        // Temporary bypass.
        eState := E_IndexState.Complete;


    E_IndexState.WaitingSupportExtended:

        (*
        bSupportExtendRequest := TRUE;

        IF bSupportExtended
            AND bTableReady
            AND bTableLocked
        THEN

            IF bManualMoveActive
                OR bPositionRecoveryActive
            THEN
                eState := E_IndexState.Complete;
            ELSE
                eState := E_IndexState.ProcessPositionReady;
            END_IF

        ELSIF tonStateTimeout.Q THEN

            eFault := E_IndexFault.SupportExtendTimeout;
            eState := E_IndexState.Fault;

        END_IF
        *)

        // Temporary bypass.
        eState := E_IndexState.Complete;


    // =====================================================
    // AUTOMATIC-CYCLE STATES
    // CURRENTLY RETAINED BUT NOT USED BY MANUAL MOVEMENT
    // =====================================================

    E_IndexState.ProcessPositionReady:

        (*
        bSupportExtendRequest := TRUE;
        *)

        IF bReleaseProcessPosition THEN

            bReleaseProcessPosition := FALSE;
            eState := E_IndexState.WaitingOperatorExchange;

        END_IF


    E_IndexState.WaitingOperatorExchange:

        (*
        bSupportExtendRequest := TRUE;
        *)

        IF bOperatorExchangeDone THEN

            bOperatorExchangeDone := FALSE;
            eState := E_IndexState.Complete;

        END_IF


    // =====================================================
    // COMPLETE
    // =====================================================

    E_IndexState.Complete:

        bDonePulse := TRUE;

        bManualMoveActive := FALSE;
        bPositionRecoveryActive := FALSE;
        bWrongPositionSupervisionActive := FALSE;

        eState := E_IndexState.Idle;


    // =====================================================
    // STOPPING
    // =====================================================

    E_IndexState.Stopping:

        // Outputs are already reset at the beginning of this method.
        IF NOT bRotatePortA THEN
            eState := E_IndexState.Idle;
        END_IF


    // =====================================================
    // FAULT
    // =====================================================

    E_IndexState.Fault:

        // No movement outputs are generated while faulted.


END_CASE


// =========================================================
// STATUS MAPPING
// =========================================================

stInternalStatus.eState := eState;
stInternalStatus.eFault := eFault;
stInternalStatus.eCurrentPosition := eCurrentPosition;

stInternalStatus.bReady :=
    eState = E_IndexState.Idle
    OR eState = E_IndexState.ProcessPositionReady;

stInternalStatus.bBusy :=
    // Support states retained for future use.
    (eState = E_IndexState.RetractingSupport)
    OR (eState = E_IndexState.WaitingSupportRetracted)

    OR (eState = E_IndexState.RotatingPortA)
    OR (eState = E_IndexState.WrongPositionRecovery)
    OR (eState = E_IndexState.StoppingPortB)
    OR (eState = E_IndexState.VerifyingPosition)

    // Support states retained for future use.
    OR (eState = E_IndexState.ExtendingSupport)
    OR (eState = E_IndexState.WaitingSupportExtended);

stInternalStatus.bFaulted :=
    eState = E_IndexState.Fault;

stInternalStatus.bDonePulse :=
    bDonePulse;

stInternalStatus.bManualMoveActive :=
    bManualMoveActive;

stInternalStatus.bPositionRecoveryActive :=
    bPositionRecoveryActive;
	
stInternalStatus.bSamePositionDetected :=
    bSamePositionDetected;

stInternalStatus.bWrongPositionTimerActive :=
    bWrongPositionSupervisionActive;

stInternalStatus.bTwoHandRequired :=
    bRequestPending
    OR (
        stInternalStatus.bBusy
        AND NOT bTableLocked
    );

stInternalStatus.bProcessPositionReady :=
    eState = E_IndexState.ProcessPositionReady;

stInternalStatus.bWaitingOperatorExchange :=
    eState = E_IndexState.WaitingOperatorExchange;


// Support feedback remains published for diagnostics, even though it
// is not currently used to permit the movement.
stInternalStatus.bSupportRetracted :=
    bSupportRetracted;

stInternalStatus.bSupportExtended :=
    bSupportExtended;

stInternalStatus.bTableReady :=
    bTableReady;

stInternalStatus.bTableLocked :=
    bTableLocked;
END_METHOD

METHOD PUBLIC GetFault : E_IndexFault
GetFault := eFault;
END_METHOD

METHOD PUBLIC GetState : E_IndexState
GetState := eState;
END_METHOD

METHOD PUBLIC GetStatus : ST_IndexStatus
GetStatus := stInternalStatus;
END_METHOD

METHOD PUBLIC IsDone : BOOL
IsDone := bDonePulse;
END_METHOD

METHOD PUBLIC IsFaulted : BOOL
IsFaulted := eState = E_IndexState.Fault;
END_METHOD

METHOD PUBLIC IsProcessPositionReady : BOOL
IsProcessPositionReady := eState = E_IndexState.ProcessPositionReady;
END_METHOD

METHOD PUBLIC IsReady : BOOL
IsReady := eState = E_IndexState.Idle OR eState = E_IndexState.ProcessPositionReady;
END_METHOD

METHOD PUBLIC ReleaseProcessPosition
IF eState = E_IndexState.ProcessPositionReady THEN bReleaseProcessPosition := TRUE; END_IF
END_METHOD

METHOD PUBLIC RequestManualMove : BOOL
RequestManualMove := FALSE;
IF eState = E_IndexState.Idle AND NOT bRequestPending THEN
    bRequestPending := TRUE;
    bManualMoveActive := TRUE;
    RequestManualMove := TRUE;
END_IF
END_METHOD

METHOD PUBLIC RequestMove : BOOL
RequestMove := FALSE;
IF eState = E_IndexState.Idle AND NOT bRequestPending THEN
    bRequestPending := TRUE;
    bManualMoveActive := FALSE;
    RequestMove := TRUE;
END_IF
END_METHOD

METHOD PUBLIC RequestPositionRecovery : BOOL
RequestPositionRecovery := FALSE;
IF eState = E_IndexState.Idle
   AND NOT bRequestPending
   AND stInternalStatus.eCurrentPosition = E_TablePosition.Unknown
THEN
    bRequestPending := TRUE;
    bManualMoveActive := FALSE;
    bPositionRecoveryActive := TRUE;
    RequestPositionRecovery := TRUE;
END_IF
END_METHOD

METHOD PUBLIC Reset
bRequestPending := FALSE;
bManualMoveActive := FALSE;
bPositionRecoveryActive := FALSE;
bWrongPositionSupervisionActive := FALSE;
bReleaseProcessPosition := FALSE;
bOperatorExchangeDone := FALSE;
eFault := E_IndexFault.None;
eState := E_IndexState.Initialising;
END_METHOD

END_FUNCTION_BLOCK

// ---- POUs/02_Components/Door/FB_MainDoorLock.TcPOU
FUNCTION_BLOCK FB_MainDoorLock
VAR
    eState           : E_MainDoorLockState := E_MainDoorLockState.Disabled;
    eFault           : E_MainDoorLockFault := E_MainDoorLockFault.None;
    stStatusInternal : ST_MainDoorLockStatus;
    tonTransition    : TON;
END_VAR

METHOD PUBLIC Cyclic : BOOL
VAR_INPUT
    bEnableAutomatic       : BOOL;
    bManualEnable          : BOOL;
    bManualLockRequest     : BOOL;
    bManualUnlockRequest   : BOOL;
    bStopRequest           : BOOL;
    bResetRequest          : BOOL;
    bDoorClosed            : BOOL;
    bDoorLocked            : BOOL;
    bIndexBusy             : BOOL;
    bProcessSafePosition   : BOOL;
    tLockTimeout           : TIME;
    tUnlockTimeout         : TIME;
	bDoorUnsafe 		   : BOOL;
END_VAR
VAR_OUTPUT
    bLockOutput            : BOOL;
	
END_VAR
// -----------------------------------------------------------------------------
// Unlock permissive
// -----------------------------------------------------------------------------
stStatusInternal.bUnlockPermissive :=
    NOT bIndexBusy
    AND bProcessSafePosition;


// -----------------------------------------------------------------------------
// This FB only supervises the main door.
//
// The physical locking is performed externally by the pneumatic system and
// TwinSAFE. This FB does not command the door lock.
// -----------------------------------------------------------------------------
bLockOutput := FALSE;


// -----------------------------------------------------------------------------
// Fault reset
// -----------------------------------------------------------------------------
IF bResetRequest THEN

    // The fault cannot be reset while TwinSAFE still reports the door unsafe.
    IF NOT bDoorUnsafe THEN

        eFault := E_MainDoorLockFault.None;

        // Restore the internal state according to the current feedbacks.
        IF bDoorClosed AND bDoorLocked THEN
            eState := E_MainDoorLockState.Locked;
        ELSE
            eState := E_MainDoorLockState.Unlocked;
        END_IF

    END_IF

END_IF


// -----------------------------------------------------------------------------
// Unsafe door condition reported by TwinSAFE
//
// Example:
//     Door not confirmed closed AND lock feedback active.
// -----------------------------------------------------------------------------
IF bDoorUnsafe THEN

    eFault := E_MainDoorLockFault.FeedbackMismatch;
    eState := E_MainDoorLockState.Fault;

END_IF


// -----------------------------------------------------------------------------
// Main door supervision state machine
// -----------------------------------------------------------------------------
CASE eState OF

    // -------------------------------------------------------------------------
    // Disabled
    // -------------------------------------------------------------------------
    E_MainDoorLockState.Disabled:

        IF bEnableAutomatic OR bManualEnable THEN

            IF bDoorClosed
                AND bDoorLocked
                AND NOT bDoorUnsafe
            THEN
                eState := E_MainDoorLockState.Locked;
            ELSE
                eState := E_MainDoorLockState.Unlocked;
            END_IF

        END_IF


    // -------------------------------------------------------------------------
    // Unlocked
    //
    // Wait for the operator to close the door.
    // An open door is not considered a fault in this state.
    // -------------------------------------------------------------------------
    E_MainDoorLockState.Unlocked:

        IF bEnableAutomatic
            OR (bManualEnable AND bManualLockRequest)
        THEN

            IF bDoorClosed AND NOT bDoorUnsafe THEN
                eState := E_MainDoorLockState.Locking;
            END_IF

        END_IF


    // -------------------------------------------------------------------------
    // Locking
    //
    // TwinSAFE and the pneumatic system perform the physical locking.
    // This FB only waits for the safe locked feedback.
    // -------------------------------------------------------------------------
    E_MainDoorLockState.Locking:

        IF bDoorUnsafe THEN

            eFault := E_MainDoorLockFault.FeedbackMismatch;
            eState := E_MainDoorLockState.Fault;

        ELSIF NOT bDoorClosed THEN

            // The door was opened before locking was confirmed.
            // Return to Unlocked without generating a fault.
            eState := E_MainDoorLockState.Unlocked;

        ELSIF bDoorLocked THEN

            eState := E_MainDoorLockState.Locked;

        ELSIF tonTransition.Q THEN

            eFault := E_MainDoorLockFault.LockTimeout;
            eState := E_MainDoorLockState.Fault;

        END_IF


    // -------------------------------------------------------------------------
    // Locked
    // -------------------------------------------------------------------------
    E_MainDoorLockState.Locked:

		// Door feedback inconsistency reported by TwinSAFE.
		IF bDoorUnsafe THEN
	
			eFault := E_MainDoorLockFault.FeedbackMismatch;
			eState := E_MainDoorLockState.Fault;
	
	
		// While automatic locking is required, the door must remain
		// physically closed and locked.
		ELSIF bEnableAutomatic
			AND (
				NOT bDoorClosed
				OR NOT bDoorLocked
			)
		THEN
	
			eFault := E_MainDoorLockFault.FeedbackMismatch;
			eState := E_MainDoorLockState.Fault;
	
	
		// Existing controlled unlock paths remain below.
		ELSIF NOT bEnableAutomatic
			AND bManualEnable
			AND bManualUnlockRequest
			AND stStatusInternal.bUnlockPermissive
		THEN
	
			eState := E_MainDoorLockState.Unlocking;
	
	
		ELSIF NOT bEnableAutomatic
			AND NOT bManualEnable
			AND bStopRequest
			AND stStatusInternal.bUnlockPermissive
		THEN
	
			eState := E_MainDoorLockState.Unlocking;
	
		END_IF


    // -------------------------------------------------------------------------
    // Unlocking
    //
    // The external safety/pneumatic system removes the locking condition.
    // This FB only waits for the lock feedback to disappear.
    // -------------------------------------------------------------------------
    E_MainDoorLockState.Unlocking:

        IF bDoorUnsafe THEN

            eFault := E_MainDoorLockFault.FeedbackMismatch;
            eState := E_MainDoorLockState.Fault;

        ELSIF NOT bDoorLocked THEN

            eState := E_MainDoorLockState.Unlocked;

        ELSIF tonTransition.Q THEN

            eFault := E_MainDoorLockFault.UnlockTimeout;
            eState := E_MainDoorLockState.Fault;

        END_IF


    // -------------------------------------------------------------------------
    // Fault
    // -------------------------------------------------------------------------
    E_MainDoorLockState.Fault:

        // No physical output is controlled by this FB.
        //
        // Recovery requires:
        //   - bDoorUnsafe = FALSE
        //   - bResetRequest = TRUE


    // -------------------------------------------------------------------------
    // Invalid internal state
    // -------------------------------------------------------------------------
    ELSE

        eFault := E_MainDoorLockFault.FeedbackMismatch;
        eState := E_MainDoorLockState.Fault;

END_CASE


// -----------------------------------------------------------------------------
// Transition timer
//
// TwinCAT SEL:
//   G = FALSE -> first value
//   G = TRUE  -> second value
//
// Locking:
//   eState = Locking -> TRUE -> tLockTimeout
//
// Unlocking:
//   eState = Locking -> FALSE -> tUnlockTimeout
// -----------------------------------------------------------------------------
tonTransition(
    IN :=
        (eState = E_MainDoorLockState.Locking)
        OR (eState = E_MainDoorLockState.Unlocking),

    PT := SEL(
        eState = E_MainDoorLockState.Locking,
        tUnlockTimeout,
        tLockTimeout
    )
);

// -----------------------------------------------------------------------------
// Status mapping
// -----------------------------------------------------------------------------
stStatusInternal.eState := eState;
stStatusInternal.eFault := eFault;

stStatusInternal.bDoorClosed := bDoorClosed;
stStatusInternal.bDoorLocked := bDoorLocked;
stStatusInternal.bDoorUnsafe := bDoorUnsafe;


// This indicates that the machine expects the door to be locked.
// It does not command the physical locking mechanism.
stStatusInternal.bLockRequest :=
    bEnableAutomatic
    OR (bManualEnable AND bManualLockRequest);


// Retained only for interface compatibility.
// This FB no longer controls a physical output.
stStatusInternal.bLockOutput := FALSE;


// Door ready for automatic operation
stStatusInternal.bReadyForAutomatic :=
    bEnableAutomatic
    AND bDoorClosed
    AND bDoorLocked
    AND NOT bDoorUnsafe
    AND (eState = E_MainDoorLockState.Locked);


stStatusInternal.bFaulted :=
    eState = E_MainDoorLockState.Fault;


// -----------------------------------------------------------------------------
// Diagnostic message
// -----------------------------------------------------------------------------
IF bDoorUnsafe THEN

    stStatusInternal.sMessage :=
        'Unsafe main door feedback';

ELSE

    CASE eState OF

        E_MainDoorLockState.Disabled:
            stStatusInternal.sMessage :=
                'Main door supervision disabled';

        E_MainDoorLockState.Unlocked:
            stStatusInternal.sMessage :=
                'Waiting for main door to close';

        E_MainDoorLockState.Locking:
            stStatusInternal.sMessage :=
                'Waiting for main door lock feedback';

        E_MainDoorLockState.Locked:
            stStatusInternal.sMessage :=
                'Main door closed and locked';

        E_MainDoorLockState.Unlocking:
            stStatusInternal.sMessage :=
                'Waiting for main door to unlock';

        E_MainDoorLockState.Fault:
            stStatusInternal.sMessage :=
                'Main door supervision fault';

        ELSE
            stStatusInternal.sMessage :=
                'Invalid main door state';

    END_CASE

END_IF


// -----------------------------------------------------------------------------
// Method result
// -----------------------------------------------------------------------------
Cyclic := NOT stStatusInternal.bFaulted;
END_METHOD

METHOD PUBLIC GetStatus : ST_MainDoorLockStatus
GetStatus := stStatusInternal;
END_METHOD

METHOD PUBLIC Initialise
eFault := E_MainDoorLockFault.None;
IF stStatusInternal.bDoorLocked THEN eState := E_MainDoorLockState.Locked; ELSE eState := E_MainDoorLockState.Unlocked; END_IF
tonTransition(IN := FALSE);
END_METHOD

METHOD PUBLIC IsFaulted : BOOL
IsFaulted := stStatusInternal.bFaulted;
END_METHOD

METHOD PUBLIC IsReadyForAutomatic : BOOL
IsReadyForAutomatic := stStatusInternal.bReadyForAutomatic;
END_METHOD

END_FUNCTION_BLOCK

// ---- POUs/02_Components/Index/FB_NestTableManager.TcPOU
FUNCTION_BLOCK FB_NestTableManager
VAR
    aNestInternal           : ARRAY[1..4] OF ST_Nest;
    aNestStatisticsInternal : ARRAY[1..4] OF ST_NestStatistics;
    aPositionToNest         : ARRAY[1..4] OF UINT := [1,2,3,4];
    bInitialised            : BOOL;
    i                       : INT;
    uiNest                  : UINT;
    uiMethodNestId          : UINT;
END_VAR

METHOD PUBLIC ClearOperatorNest
VAR_INPUT ePosition : E_TablePosition; END_VAR
uiMethodNestId := GetNestIdAtPosition(ePosition); IF uiMethodNestId >= 1 AND uiMethodNestId <= 4 THEN aNestInternal[uiMethodNestId].bProcessRequired := FALSE; aNestInternal[uiMethodNestId].bProcessComplete := FALSE; aNestInternal[uiMethodNestId].eDisposition := E_PartDisposition.None; aNestInternal[uiMethodNestId].bDispositionSent := FALSE; aNestInternal[uiMethodNestId].bOperatorExchangeComplete := FALSE; aNestInternal[uiMethodNestId].stPatchDispenseResult.bValid := FALSE; aNestInternal[uiMethodNestId].stHeatStakeResult.bValid := FALSE; aNestInternal[uiMethodNestId].stVisionResult.bValid := FALSE; aNestInternal[uiMethodNestId].stResult.bValid := FALSE; aNestInternal[uiMethodNestId].bStatisticsCounted := FALSE; END_IF
END_METHOD

METHOD PUBLIC Cyclic
VAR_INPUT
    bIndexStable : BOOL;
    eIndexPosition : E_TablePosition;
    eOperatorPosition : E_TablePosition;
    bPartPresent : BOOL;
    aNestEnabled : ARRAY[1..4] OF BOOL;
END_VAR
IF NOT bInitialised THEN
    FOR i := 1 TO 4 DO
        aNestInternal[i].nId := INT_TO_UINT(i);
        aNestStatisticsInternal[i].uiNestId := INT_TO_UINT(i);
    END_FOR
    bInitialised := TRUE;
END_IF
FOR i := 1 TO 4 DO aNestInternal[i].bEnabled := aNestEnabled[i]; END_FOR
IF bIndexStable AND (eIndexPosition <> E_TablePosition.Unknown) THEN
    CASE eIndexPosition OF
        E_TablePosition.Position1:
            aPositionToNest[1] := 1;
            aPositionToNest[2] := 4;
            aPositionToNest[3] := 3;
            aPositionToNest[4] := 2;
        E_TablePosition.Position2:
            aPositionToNest[1] := 2;
            aPositionToNest[2] := 1;
            aPositionToNest[3] := 4;
            aPositionToNest[4] := 3;
        E_TablePosition.Position3:
            aPositionToNest[1] := 3;
            aPositionToNest[2] := 2;
            aPositionToNest[3] := 1;
            aPositionToNest[4] := 4;
        E_TablePosition.Position4:
            aPositionToNest[1] := 4;
            aPositionToNest[2] := 3;
            aPositionToNest[3] := 2;
            aPositionToNest[4] := 1;
    END_CASE
    FOR i := 1 TO 4 DO
        aNestInternal[aPositionToNest[i]].ePosition := UINT_TO_E_TablePosition(INT_TO_UINT(i));
        aNestInternal[i].bPartLoadedPulse := FALSE;
        aNestInternal[i].bPartRemovedPulse := FALSE;
    END_FOR
    uiNest := aPositionToNest[TO_UINT(eOperatorPosition)];
    aNestInternal[uiNest].bPartLoadedPulse := bPartPresent AND NOT aNestInternal[uiNest].bPreviousPartPresent;
    aNestInternal[uiNest].bPartRemovedPulse := NOT bPartPresent AND aNestInternal[uiNest].bPreviousPartPresent;
    aNestInternal[uiNest].bPreviousPartPresent := bPartPresent;
    aNestInternal[uiNest].bPartPresent := bPartPresent;
END_IF
END_METHOD

METHOD PUBLIC GetAllNests : ARRAY[1..4] OF ST_Nest
GetAllNests := aNestInternal;
END_METHOD

METHOD PUBLIC GetAllNestStatistics : ARRAY[1..4] OF ST_NestStatistics
GetAllNestStatistics := aNestStatisticsInternal;
END_METHOD

METHOD PUBLIC GetNestAtPosition : ST_Nest
VAR_INPUT ePosition : E_TablePosition; END_VAR
uiMethodNestId := GetNestIdAtPosition(ePosition); IF uiMethodNestId >= 1 AND uiMethodNestId <= 4 THEN GetNestAtPosition := aNestInternal[uiMethodNestId]; END_IF
END_METHOD

METHOD PUBLIC GetNestIdAtPosition : UINT
VAR_INPUT ePosition : E_TablePosition; END_VAR
IF ePosition >= E_TablePosition.Position1 AND ePosition <= E_TablePosition.Position4 THEN GetNestIdAtPosition := aPositionToNest[TO_UINT(ePosition)]; ELSE GetNestIdAtPosition := 0; END_IF
END_METHOD

END_FUNCTION_BLOCK

// ---- POUs/03_Stations/Operator/FB_OperatorStation.TcPOU
FUNCTION_BLOCK FB_OperatorStation
VAR
    eState : E_OperatorExchangeState := E_OperatorExchangeState.Idle;
    eInstruction : E_OperatorInstruction := E_OperatorInstruction.None;
    stStatusInternal : ST_OperatorStationStatus;
    bExchangeComplete : BOOL;
END_VAR

METHOD PUBLIC Cyclic
VAR_INPUT
    bAutomaticActive : BOOL;
    bIndexStable : BOOL;
    stOperatorNest : ST_Nest;
    bPartPresent : BOOL;
    bRejectChutePartPresent : BOOL;
    bRequireRejectConfirm : BOOL;
    bAllowEmptyNestIndex : BOOL;
END_VAR
bExchangeComplete := FALSE;
IF NOT bAutomaticActive OR NOT bIndexStable THEN
    eState := E_OperatorExchangeState.Idle;
    eInstruction := E_OperatorInstruction.TableIndexing;
ELSIF stOperatorNest.stResult.bValid AND NOT stOperatorNest.stResult.bPassed THEN
    eState := E_OperatorExchangeState.WaitingForPartRemoval;
    eInstruction := E_OperatorInstruction.RemoveFailedPart;
    bExchangeComplete := NOT bPartPresent AND ((NOT bRequireRejectConfirm) OR bRejectChutePartPresent);
ELSIF stOperatorNest.stResult.bValid AND stOperatorNest.stResult.bPassed THEN
    eState := E_OperatorExchangeState.WaitingForPartRemoval;
    eInstruction := E_OperatorInstruction.RemovePassedPart;
    bExchangeComplete := NOT bPartPresent;
ELSIF bPartPresent THEN
    eState := E_OperatorExchangeState.ExchangeComplete;
    eInstruction := E_OperatorInstruction.ReadyToIndex;
    bExchangeComplete := TRUE;
ELSIF bAllowEmptyNestIndex THEN
    eState := E_OperatorExchangeState.ExchangeComplete;
    eInstruction := E_OperatorInstruction.ReadyToIndexEmpty;
    bExchangeComplete := TRUE;
ELSE
    eState := E_OperatorExchangeState.WaitingForPartLoading;
    eInstruction := E_OperatorInstruction.LoadPart;
END_IF
stStatusInternal.eState := eState;
stStatusInternal.eInstruction := eInstruction;
stStatusInternal.bExchangeComplete := bExchangeComplete;
stStatusInternal.bIndexPermissive := bExchangeComplete;
stStatusInternal.bPartPresent := bPartPresent;
stStatusInternal.bRejectChutePartPresent := bRejectChutePartPresent;
stStatusInternal.bResultValid := stOperatorNest.stResult.bValid;
stStatusInternal.bResultPassed := stOperatorNest.stResult.bPassed;
END_METHOD

METHOD PUBLIC GetInstruction : E_OperatorInstruction
GetInstruction := eInstruction;
END_METHOD

METHOD PUBLIC GetState : E_OperatorExchangeState
GetState := eState;
END_METHOD

METHOD PUBLIC GetStatus : ST_OperatorStationStatus
GetStatus := stStatusInternal;
END_METHOD

METHOD PUBLIC IndexPermissive : BOOL
IndexPermissive := stStatusInternal.bIndexPermissive;
END_METHOD

METHOD PUBLIC IsComplete : BOOL
IsComplete := bExchangeComplete;
END_METHOD

END_FUNCTION_BLOCK

// ---- POUs/03_Stations/PatchDispense/FB_PatchDispenseStation.TcPOU
FUNCTION_BLOCK FB_PatchDispenseStation
VAR
    // Method-visible diagnostics are kept at FB scope intentionally.
    eStateInternal      : E_PatchStationState := E_PatchStationState.Disabled;
    bHomeInternal       : BOOL;
    bReadyInternal      : BOOL;
    bBusyInternal       : BOOL;
    bCompleteInternal   : BOOL;
    bFaultInternal      : BOOL;
    sDiagnosticInternal : STRING(120);
END_VAR

METHOD PUBLIC Cyclic
VAR_INPUT
    bEnable       : BOOL;
    bCommissioned : BOOL;
    bStart        : BOOL;
    bReset        : BOOL;
    bSafetyOk     : BOOL;
END_VAR
VAR_OUTPUT
    stStatus      : ST_PatchStageStatus;
END_VAR
// Patch dispense foundation shell.
// No actuator is commanded until the mechanical sequence has been commissioned.
bHomeInternal := FALSE;
bReadyInternal := FALSE;
bBusyInternal := FALSE;
bCompleteInternal := FALSE;
bFaultInternal := FALSE;

IF NOT bCommissioned THEN
    eStateInternal := E_PatchStationState.Disabled;
    sDiagnosticInternal := 'Not commissioned - process sequence intentionally disabled';
ELSIF NOT bEnable OR NOT bSafetyOk THEN
    eStateInternal := E_PatchStationState.Disabled;
    sDiagnosticInternal := 'Disabled by machine state / safety';
ELSE
    // Mechanical sequence to be implemented from released design and commissioning tests.
    eStateInternal := E_PatchStationState.Homing;
    sDiagnosticInternal := 'Commissioning required - homing sequence not implemented';
END_IF

stStatus.eState := eStateInternal;
stStatus.bCommissioned := bCommissioned;
stStatus.bHome := bHomeInternal;
stStatus.bReady := bReadyInternal;
stStatus.bBusy := bBusyInternal;
stStatus.bComplete := bCompleteInternal;
stStatus.bFault := bFaultInternal;
stStatus.sDiagnostic := sDiagnosticInternal;
END_METHOD

METHOD PUBLIC Initialise
eStateInternal := E_PatchStationState.Disabled;
bHomeInternal := FALSE;
bReadyInternal := FALSE;
bBusyInternal := FALSE;
bCompleteInternal := FALSE;
bFaultInternal := FALSE;
sDiagnosticInternal := '';
END_METHOD

END_FUNCTION_BLOCK

// ---- POUs/03_Stations/HeatStake/FB_HeatStakeStation.TcPOU
FUNCTION_BLOCK FB_HeatStakeStation
VAR
    // Method-visible diagnostics are kept at FB scope intentionally.
    eStateInternal      : E_PatchStationState := E_PatchStationState.Disabled;
    bHomeInternal       : BOOL;
    bReadyInternal      : BOOL;
    bBusyInternal       : BOOL;
    bCompleteInternal   : BOOL;
    bFaultInternal      : BOOL;
    sDiagnosticInternal : STRING(120);
END_VAR

METHOD PUBLIC Cyclic
VAR_INPUT
    bEnable       : BOOL;
    bCommissioned : BOOL;
    bStart        : BOOL;
    bReset        : BOOL;
    bSafetyOk     : BOOL;
END_VAR
VAR_OUTPUT
    stStatus      : ST_PatchStageStatus;
END_VAR
// Heat stake foundation shell.
// No actuator is commanded until the mechanical sequence has been commissioned.
bHomeInternal := FALSE;
bReadyInternal := FALSE;
bBusyInternal := FALSE;
bCompleteInternal := FALSE;
bFaultInternal := FALSE;

IF NOT bCommissioned THEN
    eStateInternal := E_PatchStationState.Disabled;
    sDiagnosticInternal := 'Not commissioned - process sequence intentionally disabled';
ELSIF NOT bEnable OR NOT bSafetyOk THEN
    eStateInternal := E_PatchStationState.Disabled;
    sDiagnosticInternal := 'Disabled by machine state / safety';
ELSE
    // Mechanical sequence to be implemented from released design and commissioning tests.
    eStateInternal := E_PatchStationState.Homing;
    sDiagnosticInternal := 'Commissioning required - homing sequence not implemented';
END_IF

stStatus.eState := eStateInternal;
stStatus.bCommissioned := bCommissioned;
stStatus.bHome := bHomeInternal;
stStatus.bReady := bReadyInternal;
stStatus.bBusy := bBusyInternal;
stStatus.bComplete := bCompleteInternal;
stStatus.bFault := bFaultInternal;
stStatus.sDiagnostic := sDiagnosticInternal;
END_METHOD

METHOD PUBLIC Initialise
eStateInternal := E_PatchStationState.Disabled;
bHomeInternal := FALSE;
bReadyInternal := FALSE;
bBusyInternal := FALSE;
bCompleteInternal := FALSE;
bFaultInternal := FALSE;
sDiagnosticInternal := '';
END_METHOD

END_FUNCTION_BLOCK

// ---- POUs/03_Stations/Vision/FB_VisionStation.TcPOU
FUNCTION_BLOCK FB_VisionStation
VAR
    // Method-visible diagnostics are kept at FB scope intentionally.
    eStateInternal      : E_PatchStationState := E_PatchStationState.Disabled;
    bHomeInternal       : BOOL;
    bReadyInternal      : BOOL;
    bBusyInternal       : BOOL;
    bCompleteInternal   : BOOL;
    bFaultInternal      : BOOL;
    sDiagnosticInternal : STRING(120);
END_VAR

METHOD PUBLIC Cyclic
VAR_INPUT
    bEnable       : BOOL;
    bCommissioned : BOOL;
    bStart        : BOOL;
    bReset        : BOOL;
    bSafetyOk     : BOOL;
END_VAR
VAR_OUTPUT
    stStatus      : ST_PatchStageStatus;
END_VAR
// Vision inspection foundation shell.
// No actuator is commanded until the mechanical sequence has been commissioned.
bHomeInternal := FALSE;
bReadyInternal := FALSE;
bBusyInternal := FALSE;
bCompleteInternal := FALSE;
bFaultInternal := FALSE;

IF NOT bCommissioned THEN
    eStateInternal := E_PatchStationState.Disabled;
    sDiagnosticInternal := 'Not commissioned - process sequence intentionally disabled';
ELSIF NOT bEnable OR NOT bSafetyOk THEN
    eStateInternal := E_PatchStationState.Disabled;
    sDiagnosticInternal := 'Disabled by machine state / safety';
ELSE
    // Mechanical sequence to be implemented from released design and commissioning tests.
    eStateInternal := E_PatchStationState.Homing;
    sDiagnosticInternal := 'Commissioning required - homing sequence not implemented';
END_IF

stStatus.eState := eStateInternal;
stStatus.bCommissioned := bCommissioned;
stStatus.bHome := bHomeInternal;
stStatus.bReady := bReadyInternal;
stStatus.bBusy := bBusyInternal;
stStatus.bComplete := bCompleteInternal;
stStatus.bFault := bFaultInternal;
stStatus.sDiagnostic := sDiagnosticInternal;
END_METHOD

METHOD PUBLIC Initialise
eStateInternal := E_PatchStationState.Disabled;
bHomeInternal := FALSE;
bReadyInternal := FALSE;
bBusyInternal := FALSE;
bCompleteInternal := FALSE;
bFaultInternal := FALSE;
sDiagnosticInternal := '';
END_METHOD

END_FUNCTION_BLOCK

// ---- POUs/01_Core/Machine/FB_PatchPressCommissioningGuard.TcPOU
FUNCTION_BLOCK FB_PatchPressCommissioningGuard
VAR
    // Deliberately at FB scope so values remain visible online while debugging.
    bAllStationsCommissionedInternal : BOOL;
    bAutoCycleAllowedInternal        : BOOL;
    sBlockReasonInternal             : STRING(160);
END_VAR

METHOD PUBLIC Cyclic
VAR_INPUT
    bDispenseCommissioned : BOOL;
    bHeatStakeCommissioned: BOOL;
    bVisionCommissioned   : BOOL;
    bCoreCommissioningMode: BOOL;
    bCoreReady            : BOOL;
END_VAR
VAR_OUTPUT
    bAutoCycleAllowed     : BOOL;
    sBlockReason          : STRING(160);
END_VAR
bAllStationsCommissionedInternal := bDispenseCommissioned AND bHeatStakeCommissioned AND bVisionCommissioned;
bAutoCycleAllowedInternal := bCoreReady AND (bAllStationsCommissionedInternal OR bCoreCommissioningMode);

IF NOT bCoreReady THEN
    sBlockReasonInternal := 'Core machine not ready';
ELSIF bCoreCommissioningMode THEN
    sBlockReasonInternal := '';
ELSIF NOT bDispenseCommissioned THEN
    sBlockReasonInternal := 'Patch dispense station not commissioned';
ELSIF NOT bHeatStakeCommissioned THEN
    sBlockReasonInternal := 'Heat stake station not commissioned';
ELSIF NOT bVisionCommissioned THEN
    sBlockReasonInternal := 'Vision station not commissioned';
ELSE
    sBlockReasonInternal := '';
END_IF

bAutoCycleAllowed := bAutoCycleAllowedInternal;
sBlockReason := sBlockReasonInternal;
END_METHOD

END_FUNCTION_BLOCK

// ---- POUs/05_AlarmsAndEvents/PRG_Events.TcPOU
PROGRAM PRG_Events
VAR
    fbEventsManager : FB_EventsManager;
    tonUpSupplyLost : TON;
    tonUsSupplyLost : TON;
    ton48VSupplyLost : TON;
    tonIndexPositionInvalid : TON;
END_VAR

GVL_MASTER.sSystemDate := '';
GVL_MASTER.sSystemTime := '';
GVL_MASTER.stStationEvents[0].aEvents[0].bFault := TRUE;
GVL_MASTER.stStationEvents[0].aEvents[0].bEventFlag := NOT GVL_MASTER.stInputs.bEmergencyStopChannel1 OR NOT GVL_MASTER.stInputs.bEmergencyStopChannel2;
GVL_MASTER.stStationEvents[0].aEvents[0].bEventText := 'E-stop activated';
GVL_MASTER.stStationEvents[0].aEvents[0].sSolution := 'Release E-stop and reset Safety';
GVL_MASTER.stStationEvents[0].aEvents[1].bFault := TRUE;
GVL_MASTER.stStationEvents[0].aEvents[1].bEventFlag := NOT GVL_MASTER.stInputs.bMainDoorChannel1 OR NOT GVL_MASTER.stInputs.bMainDoorChannel2;
GVL_MASTER.stStationEvents[0].aEvents[1].bEventText := 'Main door safety circuit open';
GVL_MASTER.stStationEvents[0].aEvents[1].sSolution := 'Close main door and reset Safety';
GVL_MASTER.stStationEvents[0].aEvents[2].bFault := TRUE;
GVL_MASTER.stStationEvents[0].aEvents[2].bEventFlag := (NOT GVL_MASTER.stInputs.bLeftFlapChannel1 OR NOT GVL_MASTER.stInputs.bLeftFlapChannel2) AND (GVL_MASTER.stStatus.eMachineState <> E_MachineState.PowerUp);
GVL_MASTER.stStationEvents[0].aEvents[2].bEventText := 'Left safety flap active';
GVL_MASTER.stStationEvents[0].aEvents[2].sSolution := 'Clear left flap and reset Safety';
GVL_MASTER.stStationEvents[0].aEvents[3].bFault := TRUE;
GVL_MASTER.stStationEvents[0].aEvents[3].bEventFlag := (NOT GVL_MASTER.stInputs.bRightFlapChannel1 OR NOT GVL_MASTER.stInputs.bRightFlapChannel2) AND (GVL_MASTER.stStatus.eMachineState <> E_MachineState.PowerUp);
GVL_MASTER.stStationEvents[0].aEvents[3].bEventText := 'Right safety flap active';
GVL_MASTER.stStationEvents[0].aEvents[3].sSolution := 'Clear right flap and reset Safety';
GVL_MASTER.stStationEvents[0].aEvents[4].bCycleStopRequest := TRUE;
GVL_MASTER.stStationEvents[0].aEvents[4].bEventFlag := GVL_MASTER.stCommand.bStop;
GVL_MASTER.stStationEvents[0].aEvents[4].bEventText := 'Cycle stop requested';
GVL_MASTER.stStationEvents[0].aEvents[4].sSolution := 'Wait for cycle to stop';
GVL_MASTER.stStationEvents[0].aEvents[5].bFault := TRUE;
GVL_MASTER.stStationEvents[0].aEvents[5].bEventFlag := GVL_MASTER.stStatus.bInitialisationTimeoutFault;
GVL_MASTER.stStationEvents[0].aEvents[5].bEventText := 'System initialisation timeout';
GVL_MASTER.stStationEvents[0].aEvents[5].sSolution := 'Check initialisation conditions';
GVL_MASTER.stStationEvents[0].aEvents[6].bFault := TRUE;
GVL_MASTER.stStationEvents[0].aEvents[6].bEventFlag := GVL_MASTER.stStatus.bStoppingTimeoutFault;
GVL_MASTER.stStationEvents[0].aEvents[6].bEventText := 'System stopping timeout';
GVL_MASTER.stStationEvents[0].aEvents[6].sSolution := 'Check index and machine safe state';
tonUpSupplyLost(IN := NOT GVL_MASTER.stInputs.bUp24VPowerSupplyOk AND (GVL_MASTER.stStatus.eMachineState <> E_MachineState.PowerUp), PT := T#1S);
GVL_MASTER.stStationEvents[0].aEvents[7].bFault := TRUE;
GVL_MASTER.stStationEvents[0].aEvents[7].bEventFlag := tonUpSupplyLost.Q;
GVL_MASTER.stStationEvents[0].aEvents[7].bEventText := '24 V Up supply fault';
GVL_MASTER.stStationEvents[0].aEvents[7].sSolution := 'Check 24 V Up power supply';
tonUsSupplyLost(IN := NOT GVL_MASTER.stInputs.bUs24VPowerSupplyOk AND (GVL_MASTER.stStatus.eMachineState <> E_MachineState.PowerUp), PT := T#1S);
GVL_MASTER.stStationEvents[0].aEvents[8].bFault := TRUE;
GVL_MASTER.stStationEvents[0].aEvents[8].bEventFlag := tonUsSupplyLost.Q;
GVL_MASTER.stStationEvents[0].aEvents[8].bEventText := '24 V Us supply fault';
GVL_MASTER.stStationEvents[0].aEvents[8].sSolution := 'Check 24 V Us power supply';
ton48VSupplyLost(IN := NOT GVL_MASTER.stInputs.b48VPowerSupplyOk AND (GVL_MASTER.stStatus.eMachineState <> E_MachineState.PowerUp), PT := T#1S);
GVL_MASTER.stStationEvents[0].aEvents[9].bFault := TRUE;
GVL_MASTER.stStationEvents[0].aEvents[9].bEventFlag := ton48VSupplyLost.Q;
GVL_MASTER.stStationEvents[0].aEvents[9].bEventText := '48 V Up supply fault';
GVL_MASTER.stStationEvents[0].aEvents[9].sSolution := 'Check 48 V power supply';
tonIndexPositionInvalid(IN := GVL_MASTER.stInputs.bIndexReady AND GVL_MASTER.stInputs.bIndexLocked AND (GVL_MASTER.stInputs.eIndexPosition = E_TablePosition.Unknown), PT := T#500MS);
GVL_MASTER.stStationEvents[2].aEvents[0].bFault := TRUE;
GVL_MASTER.stStationEvents[2].aEvents[0].bEventFlag := tonIndexPositionInvalid.Q;
GVL_MASTER.stStationEvents[2].aEvents[0].bEventText := 'Index position sensors invalid';
GVL_MASTER.stStationEvents[2].aEvents[0].sSolution := 'Check index position sensors';
GVL_MASTER.stStationEvents[1].aEvents[0].bMessage := TRUE;
GVL_MASTER.stStationEvents[1].aEvents[0].bPersistentMessage := TRUE;
GVL_MASTER.stStationEvents[1].aEvents[0].bEventFlag := NOT GVL_MASTER.stStatus.bAllStationsCommissioned;
GVL_MASTER.stStationEvents[1].aEvents[0].bEventText := GVL_MASTER.stStatus.sAutoCycleBlockReason;
GVL_MASTER.stStationEvents[1].aEvents[0].sSolution := 'Commission Patch Dispense, Heat Stake and Vision stations';
fbEventsManager(bPulse := TRUE, sSystemTime := GVL_MASTER.sSystemTime, sSystemDate := GVL_MASTER.sSystemDate, bDataWritedInCSV := FALSE, nArraySize := 4, bMachineMessage := GVL_MASTER.stStatus.sMachineMessage, eMachineState := GVL_MASTER.stStatus.eMachineState, stStationEvents := GVL_MASTER.stStationEvents, stEventsAssigment := GVL_MASTER.stEventsAssigment, bResetFaults := GVL_MASTER.stCommand.bReset, bMachineFault => GVL_MASTER.bMachineFault, bCycleStopRequest => GVL_MASTER.bCycleStopRequest, astActiveEvents => GVL_MASTER.astActiveEvents, astEventsHistory => GVL_Persistent.astEventsHistory);
GVL_HMI.astActiveEvents := GVL_MASTER.astActiveEvents;
GVL_HMI.astEventsHistory := GVL_Persistent.astEventsHistory;
GVL_HMI.stEventsAssigment := GVL_MASTER.stEventsAssigment;

END_PROGRAM

// ---- POUs/05_AlarmsAndEvents/FB_EventsManager.TcPOU
FUNCTION_BLOCK FB_EventsManager
VAR_INPUT
	bPulse					: BOOL;
	sSystemTime				: STRING(255);
	sSystemDate				: STRING(255);
	bDataWritedInCSV		: BOOL;
	nArraySize				: DINT;
	bMachineMessage			: STRING;
	eMachineState 			: E_MachineState;
END_VAR
VAR_OUTPUT
    bMachineFault            : BOOL;
    bCycleStopRequest        : BOOL;
	astActiveEvents			: ARRAY [0..50] OF ST_ActiveEvents;
	astEventsHistory		: ARRAY[0..200] OF ST_EventsHistory;
END_VAR
VAR
	i								: ARRAY [0..1] OF DINT;
	j								: ARRAY [0..1] OF DINT;
	m								: ARRAY [0..3] OF DINT;
	k								: ARRAY [0..1] OF DINT;
	l								: DINT;
	n								: DINT;
	
	bEventsAssigmentSignal			: BOOL		:= TRUE;
    bStationFaultCondition   : BOOL;
    bStationStopCondition    : BOOL;
END_VAR

VAR_IN_OUT
	
	stStationEvents			: ARRAY[0..4] OF ST_StationEvents;
	stEventsAssigment		: ST_EventsAssigmentGeneral;
	bResetFaults			: BOOL;
	
END_VAR

ACT_FaultTrig();

ACT_EventTextAssigment();

ACT_ActiveEvents_DataHistory();

// Row zero is permanently reserved for the operational instruction.
astActiveEvents[0].sEventTex := bMachineMessage;
astActiveEvents[0].sType := 'Message';
astActiveEvents[0].abType := 3;
astActiveEvents[0].sSolution := '';

ACTION ACT_ActiveEvents_DataHistory:
// ============================================================================
// ACTIVE EVENTS AND EVENT HISTORY
// ============================================================================
//
// astActiveEvents[0]:
//     Reserved exclusively for the current machine message.
//
// astActiveEvents[1..50]:
//     Active Faults and Cycle Stop Requests.
//
// astEventsHistory:
//     Complete event history.
//
// EVENT BEHAVIOUR:
//
// MESSAGE:
//     - Operator instruction.
//     - Displayed only through astActiveEvents[0].
//     - Never added to rows 1..50.
//
// FAULT:
//     - Latched individually through bActive.
//     - Displayed only while the machine is in Fault.
//     - Remains latched after the live condition disappears.
//     - Cleared by Reset only after bEventFlag is FALSE.
//
// CYCLE STOP REQUEST:
//     - Latched individually through bActive.
//     - Displayed in any machine state.
//     - Remains visible after the live condition disappears.
//     - Cleared by Reset only after bEventFlag is FALSE.
//
// bEventFlag:
//     Live condition.
//
// bActive:
//     Individual event presentation latch.
//
// ============================================================================


IF bPulse THEN

    // ------------------------------------------------------------------------
    // REBUILD ACTIVE EVENT GRID
    // ------------------------------------------------------------------------
    // Row 0 is intentionally preserved because it contains the current
    // machine instruction/message.
    // ------------------------------------------------------------------------

    FOR l := 1 TO 50 DO

        astActiveEvents[l].sEventTex := '';
        astActiveEvents[l].sType := '';
        astActiveEvents[l].abType := 0;
        astActiveEvents[l].sSolution := '';

    END_FOR


    // Rows 1..50 are used for Faults and Alerts.
    l := 0;


    // ------------------------------------------------------------------------
    // SCAN ALL STATION EVENTS
    // ------------------------------------------------------------------------

    FOR k[0] := 0 TO nArraySize DO

        FOR k[1] := 0 TO 100 DO


            // =================================================================
            // FAULT
            // =================================================================

            IF stStationEvents[k[0]].aEvents[k[1]].bFault THEN


                // -------------------------------------------------------------
                // NEW FAULT DETECTED
                // -------------------------------------------------------------
                // Register in history only once, when the live condition
                // activates an event that was not already latched.
                // -------------------------------------------------------------

                IF stStationEvents[k[0]].aEvents[k[1]].bEventFlag
                    AND NOT stStationEvents[k[0]].aEvents[k[1]].bActive
                THEN

                    // Shift history.
                    FOR n := 200 TO 1 BY -1 DO

                        astEventsHistory[n] :=
                            astEventsHistory[n - 1];

                    END_FOR


                    // Insert newest event.
                    astEventsHistory[0].sEventTex :=
                        stStationEvents[k[0]].aEvents[k[1]].bEventTextHMI;

                    astEventsHistory[0].sType :=
                        'Fault';

                    astEventsHistory[0].abType :=
                        1;

                    astEventsHistory[0].sDate :=
                        sSystemDate;

                    astEventsHistory[0].sTime :=
                        sSystemTime;


                    // Latch the individual event.
                    stStationEvents[k[0]].aEvents[k[1]].bActive :=
                        TRUE;

                END_IF


                // -------------------------------------------------------------
                // RESET FAULT LATCH
                // -------------------------------------------------------------
                // Reset is allowed to clear the individual event only after
                // the originating fault condition has disappeared.
                // -------------------------------------------------------------

                IF bResetFaults
                    AND NOT stStationEvents[k[0]].aEvents[k[1]].bEventFlag
                THEN

                    stStationEvents[k[0]].aEvents[k[1]].bActive :=
                        FALSE;

                END_IF


                // -------------------------------------------------------------
                // ACTIVE GRID
                // -------------------------------------------------------------
                // Faults are shown only while the machine itself is in Fault.
                //
                // bActive allows the original cause to remain displayed after
                // bEventFlag has returned FALSE, until the operator resets.
                // -------------------------------------------------------------

                IF stStationEvents[k[0]].aEvents[k[1]].bActive
                    AND eMachineState = E_MachineState.Fault
                THEN

                    IF l < 50 THEN

                        l := l + 1;

                        astActiveEvents[l].sEventTex :=
                            stStationEvents[k[0]].aEvents[k[1]].bEventTextHMI;

                        astActiveEvents[l].sType :=
                            'Fault';

                        astActiveEvents[l].abType :=
                            1;

                        astActiveEvents[l].sSolution :=
                            stStationEvents[k[0]].aEvents[k[1]].sSolution;

                    END_IF

                END_IF



            // =================================================================
            // CYCLE STOP REQUEST / ALERT
            // =================================================================

            ELSIF stStationEvents[k[0]].aEvents[k[1]].bCycleStopRequest THEN


                // -------------------------------------------------------------
                // NEW ALERT DETECTED
                // -------------------------------------------------------------

                IF stStationEvents[k[0]].aEvents[k[1]].bEventFlag
                    AND NOT stStationEvents[k[0]].aEvents[k[1]].bActive
                THEN

                    // Shift history.
                    FOR n := 200 TO 1 BY -1 DO

                        astEventsHistory[n] :=
                            astEventsHistory[n - 1];

                    END_FOR


                    // Insert newest event.
                    astEventsHistory[0].sEventTex :=
                        stStationEvents[k[0]].aEvents[k[1]].bEventTextHMI;

                    astEventsHistory[0].sType :=
                        'Cycle Stop Request';

                    astEventsHistory[0].abType :=
                        2;

                    astEventsHistory[0].sDate :=
                        sSystemDate;

                    astEventsHistory[0].sTime :=
                        sSystemTime;


                    // Latch the individual Alert.
                    stStationEvents[k[0]].aEvents[k[1]].bActive :=
                        TRUE;

                END_IF


                // -------------------------------------------------------------
                // RESET ALERT LATCH
                // -------------------------------------------------------------
                // The Alert remains displayed after the live condition has
                // disappeared and is acknowledged by Reset.
                // -------------------------------------------------------------

                IF bResetFaults
                    AND NOT stStationEvents[k[0]].aEvents[k[1]].bEventFlag
                THEN

                    stStationEvents[k[0]].aEvents[k[1]].bActive :=
                        FALSE;

                END_IF


                // -------------------------------------------------------------
                // ACTIVE GRID
                // -------------------------------------------------------------
                // Alerts may be shown in any machine state.
                // -------------------------------------------------------------

                IF stStationEvents[k[0]].aEvents[k[1]].bActive THEN

                    IF l < 50 THEN

                        l := l + 1;

                        astActiveEvents[l].sEventTex :=
                            stStationEvents[k[0]].aEvents[k[1]].bEventTextHMI;

                        astActiveEvents[l].sType :=
                            'Cycle Stop Request';

                        astActiveEvents[l].abType :=
                            2;

                        astActiveEvents[l].sSolution :=
                            stStationEvents[k[0]].aEvents[k[1]].sSolution;

                    END_IF

                END_IF



            // =================================================================
            // MESSAGE
            // =================================================================
            //
            // Messages are instructions for the operator.
            //
            // They are NOT inserted into astActiveEvents[1..50].
            // Row 0 remains exclusively responsible for the current machine
            // instruction through sMachineMessage.
            //
            // bActive is not used as an operator-reset latch for Messages.
            // =================================================================

            ELSIF stStationEvents[k[0]].aEvents[k[1]].bMessage THEN


                // -------------------------------------------------------------
                // OPTIONAL MESSAGE HISTORY
                // -------------------------------------------------------------
                // Preserve the existing ability to register message events in
                // history, but rearm them automatically when their condition
                // disappears because Messages do not require operator Reset.
                // -------------------------------------------------------------

                IF stStationEvents[k[0]].aEvents[k[1]].bEventFlag
                    AND NOT stStationEvents[k[0]].aEvents[k[1]].bActive
                THEN

                    FOR n := 200 TO 1 BY -1 DO

                        astEventsHistory[n] :=
                            astEventsHistory[n - 1];

                    END_FOR


                    astEventsHistory[0].sEventTex :=
                        stStationEvents[k[0]].aEvents[k[1]].bEventTextHMI;

                    astEventsHistory[0].sType :=
                        'Message';

                    astEventsHistory[0].abType :=
                        3;

                    astEventsHistory[0].sDate :=
                        sSystemDate;

                    astEventsHistory[0].sTime :=
                        sSystemTime;


                    stStationEvents[k[0]].aEvents[k[1]].bActive :=
                        TRUE;

                END_IF


                // Messages automatically rearm when their live condition ends.
                IF NOT stStationEvents[k[0]].aEvents[k[1]].bEventFlag THEN

                    stStationEvents[k[0]].aEvents[k[1]].bActive :=
                        FALSE;

                END_IF

                // Live message: shown in Active Events while the condition is
                // TRUE and cannot be acknowledged/reset by the operator.
                IF stStationEvents[k[0]].aEvents[k[1]].bPersistentMessage
                    AND stStationEvents[k[0]].aEvents[k[1]].bEventFlag
                THEN

                    IF l < 50 THEN
                        l := l + 1;
                        astActiveEvents[l].sEventTex :=
                            stStationEvents[k[0]].aEvents[k[1]].bEventTextHMI;
                        astActiveEvents[l].sType := 'Message';
                        astActiveEvents[l].abType := 3;
                        astActiveEvents[l].sSolution :=
                            stStationEvents[k[0]].aEvents[k[1]].sSolution;
                    END_IF

                END_IF


            END_IF


        END_FOR

    END_FOR


END_IF
END_ACTION

ACTION ACT_EventTextAssigment:

FOR j[0] := 0 TO nArraySize DO
	
	FOR j[1] := 0 TO 100 DO 
		
		IF stStationEvents[j[0]].aEvents[j[1]].bFault THEN
			
			m[0]											:= m[0]+1;
			
			stStationEvents[j[0]].aEvents[j[1]].bEventTextHMI	:= 		CONCAT( STR1 := 'N ', STR2 := 
																CONCAT( STR1 := DINT_TO_STRING(m[0]), str2 := 
																CONCAT( STR1 :='-Station' , STR2 := 
																CONCAT( STR1 := DINT_TO_STRING(j[0]), STR2 := 
																CONCAT( STR1 :=' - ', str2 := stStationEvents[j[0]].aEvents[j[1]].bEventText )))));
			stStationEvents[j[0]].aEvents[j[1]].bAssignedID	:= 	m[0];				
			
			//EVENTS ASSIGMENT
			stEventsAssigment.astFaultEvents[m[0]].sEventText	:= stStationEvents[j[0]].aEvents[j[1]].bEventTextHMI;
			stEventsAssigment.astFaultEvents[m[0]].sSolution	:= stStationEvents[j[0]].aEvents[j[1]].sSolution;
			
		ELSIF stStationEvents[j[0]].aEvents[j[1]].bCycleStopRequest THEN
		
			m[2]											:= m[2]+1;	
			
			stStationEvents[j[0]].aEvents[j[1]].bEventTextHMI	:= 		CONCAT( STR1 := 'N ', STR2 := 
																CONCAT( STR1 := DINT_TO_STRING(m[2]), str2 := 
																CONCAT( STR1 :='-Station' , STR2 := 
																CONCAT( STR1 := DINT_TO_STRING(j[0]), STR2 := 
																CONCAT( STR1 :=' - ', str2 := stStationEvents[j[0]].aEvents[j[1]].bEventText )))));
			stStationEvents[j[0]].aEvents[j[1]].bAssignedID	:= 	m[2];													

			//EVENTS ASSIGMENT
			stEventsAssigment.astCycleStopRequestEvents[m[2]].sEventText	:= stStationEvents[j[0]].aEvents[j[1]].bEventTextHMI;
			stEventsAssigment.astCycleStopRequestEvents[m[2]].sSolution	:= stStationEvents[j[0]].aEvents[j[1]].sSolution;
			
		ELSIF stStationEvents[j[0]].aEvents[j[1]].bMessage THEN
			
			m[3]											:= m[3]+1;
			
			stStationEvents[j[0]].aEvents[j[1]].bEventTextHMI	:= 		CONCAT( STR1 := 'N ', STR2 := 
																CONCAT( STR1 := DINT_TO_STRING(m[3]), str2 := 
																CONCAT( STR1 :='-Station' , STR2 := 
																CONCAT( STR1 := DINT_TO_STRING(j[0]), STR2 := 
																CONCAT( STR1 :=' - ', str2 := stStationEvents[j[0]].aEvents[j[1]].bEventText )))));
			stStationEvents[j[0]].aEvents[j[1]].bAssignedID	:= 	m[3];													
				
			//EVENTS ASSIGMENT
			stEventsAssigment.astMessage[m[3]].sEventText	:= stStationEvents[j[0]].aEvents[j[1]].bEventTextHMI;
			stEventsAssigment.astMessage[m[3]].sSolution	:= stStationEvents[j[0]].aEvents[j[1]].sSolution;	
			
		END_IF
		
	END_FOR
	
	
END_FOR
j[0]														:= 0;
j[1]														:= 0;
m[0]														:= 0;
m[1]														:= 0;
m[2]														:= 0;
m[3]														:= 0;
END_ACTION

ACTION ACT_FaultTrig:
// Deterministic station aggregation. Classification is fixed in each point;
// bEventFlag is the live condition. Station flags are latched until Reset.
bMachineFault := FALSE;
bCycleStopRequest := FALSE;

FOR i[0] := 0 TO nArraySize DO
    bStationFaultCondition := FALSE;
    bStationStopCondition := FALSE;

    FOR i[1] := 0 TO 100 DO
        bStationFaultCondition := bStationFaultCondition
            OR (stStationEvents[i[0]].aEvents[i[1]].bFault
                AND stStationEvents[i[0]].aEvents[i[1]].bEventFlag);

        bStationStopCondition := bStationStopCondition
            OR (stStationEvents[i[0]].aEvents[i[1]].bCycleStopRequest
                AND stStationEvents[i[0]].aEvents[i[1]].bEventFlag);
    END_FOR

    IF bStationFaultCondition THEN
        stStationEvents[i[0]].bFault := TRUE;
    ELSIF bResetFaults THEN
        stStationEvents[i[0]].bFault := FALSE;
    END_IF

    IF bStationStopCondition THEN
        stStationEvents[i[0]].bCycleStopRequest := TRUE;
    ELSIF bResetFaults THEN
        stStationEvents[i[0]].bCycleStopRequest := FALSE;
    END_IF

    bMachineFault := bMachineFault OR stStationEvents[i[0]].bFault;
    bCycleStopRequest := bCycleStopRequest OR stStationEvents[i[0]].bCycleStopRequest;
END_FOR
END_ACTION

END_FUNCTION_BLOCK

// ---- POUs/00_Application/PRG_HmiStatus.TcPOU
PROGRAM PRG_HmiStatus
VAR
END_VAR

GVL_HMI.stStatus.eMachineState := GVL_MASTER.stStatus.eMachineState;
GVL_HMI.stStatus.eIndexState := GVL_MASTER.stStatus.eIndexState;
GVL_HMI.stStatus.eIndexPosition := GVL_MASTER.stInputs.eIndexPosition;
GVL_HMI.stStatus.bReady := GVL_MASTER.stStatus.bReady;
GVL_HMI.stStatus.bBusy := GVL_MASTER.stStatus.bBusy;
GVL_HMI.stStatus.bFaulted := GVL_MASTER.stStatus.bFaulted;
GVL_HMI.stStatus.bTwoHandsSafe := GVL_MASTER.stInputs.bTwoHandsSafe;
GVL_HMI.stStatus.bLoadingStationEaglePresent := GVL_MASTER.stInputs.bLoadingStationEaglePresent;
GVL_HMI.stStatus.bRejectChutePartPresent := GVL_MASTER.stInputs.bRejectChutePartPresent;
GVL_HMI.stStatus.bHeatStakeEaglePresent := GVL_MASTER.stInputs.bHeatStakeEaglePresent;
GVL_HMI.stStatus.bHeatStakePatchPresent := GVL_MASTER.stInputs.bHeatStakePatchPresent;
GVL_HMI.stStatus.bPbupMagnetPresent := GVL_MASTER.stInputs.bPbupMagnetPresent;
GVL_HMI.stStatus.bIndexReady := GVL_MASTER.stInputs.bIndexReady;
GVL_HMI.stStatus.bIndexLocked := GVL_MASTER.stInputs.bIndexLocked;
GVL_HMI.stStatus.bIndexCompletedSensor := GVL_MASTER.stInputs.bIndexCompletedSensor;
GVL_HMI.stStatus.bMainDoorClosed := GVL_MASTER.stInputs.bMainDoorClosed;
GVL_HMI.stStatus.bMainDoorLocked := GVL_MASTER.stInputs.bMainDoorLocked;
GVL_HMI.stStatus.bStartButtonActive := GVL_MASTER.stInputs.bStartButton;
GVL_HMI.stStatus.bStopButtonActive := GVL_MASTER.stInputs.bStopButton;
GVL_HMI.stStatus.bResetButtonActive := GVL_MASTER.stInputs.bResetButton;
GVL_HMI.stStatus.bStartButtonLamp := GVL_MASTER.stOutputs.bLedStart;
GVL_HMI.stStatus.bUp24VPowerSupplyOk := GVL_MASTER.stInputs.bUp24VPowerSupplyOk;
GVL_HMI.stStatus.bUs24VPowerSupplyOk := GVL_MASTER.stInputs.bUs24VPowerSupplyOk;
GVL_HMI.stStatus.b48VPowerSupplyOk := GVL_MASTER.stInputs.b48VPowerSupplyOk;
GVL_HMI.stStatus.bMainDoorDiagnosticOk := GVL_MASTER.stInputs.bMainDoorDiagnosticOk;
GVL_HMI.stStatus.bMs6FeedbackOk := GVL_MASTER.stInputs.bMs6FeedbackOk;
GVL_HMI.stStatus.bAirExhausted := GVL_MASTER.stInputs.bAirExhausted;
GVL_HMI.stStatus.bLeftFlapSafe := GVL_MASTER.stInputs.stSafety.bLeftFlapSafe;
GVL_HMI.stStatus.bRightFlapSafe := GVL_MASTER.stInputs.stSafety.bRightFlapSafe;
GVL_HMI.stStatus.bEnableSettings := GVL_MASTER.stStatus.bEnableSetting;
GVL_HMI.stStatus.bAllStationsCommissioned := GVL_MASTER.stStatus.bAllStationsCommissioned;
GVL_HMI.stStatus.bAutoCycleAllowed := GVL_MASTER.stStatus.bAutoCycleAllowed;
GVL_HMI.stStatus.stPatchDispense := GVL_MASTER.stStatus.stPatchDispense;
GVL_HMI.stStatus.stHeatStake := GVL_MASTER.stStatus.stHeatStake;
GVL_HMI.stStatus.stVision := GVL_MASTER.stStatus.stVision;
GVL_HMI.stStatus.eOperatorInstruction := GVL_MASTER.stStatus.eOperatorInstruction;
GVL_HMI.stStatus.stOperatorStation := GVL_MASTER.stStatus.stOperatorStation;
GVL_HMI.stStatus.aNest := GVL_MASTER.stStatus.aNest;
GVL_HMI.stStatus.sMachineMessage := GVL_MASTER.stStatus.sMachineMessage;
GVL_HMI.stStatus.sOperatorMessage := GVL_MASTER.stStatus.sOperatorMessage;
GVL_HMI.stStatus.sAutoCycleBlockReason := GVL_MASTER.stStatus.sAutoCycleBlockReason;
GVL_HMI.stStatistics.aNest := GVL_MASTER.stStatus.aNestStatistics;
CASE GVL_MASTER.stInputs.eIndexPosition OF
    E_TablePosition.Position1: GVL_HMI.stStatus.iNestRotationAngle := 0;
    E_TablePosition.Position2: GVL_HMI.stStatus.iNestRotationAngle := 270;
    E_TablePosition.Position3: GVL_HMI.stStatus.iNestRotationAngle := 180;
    E_TablePosition.Position4: GVL_HMI.stStatus.iNestRotationAngle := 90;
ELSE GVL_HMI.stStatus.iNestRotationAngle := 0;
END_CASE
CASE GVL_MASTER.stStatus.eMachineState OF
    E_MachineState.PowerUp: GVL_HMI.StatusHMI.sMachineStatusText := 'SYSTEM POWER UP'; GVL_HMI.StatusHMI.sBannerBckColor := GVL_HMI.sYELLOW; GVL_HMI.StatusHMI.sBannerTextColor := GVL_HMI.sBLACK;
    E_MachineState.Initialising: GVL_HMI.StatusHMI.sMachineStatusText := 'SYSTEM INITIALIZING'; GVL_HMI.StatusHMI.sBannerBckColor := GVL_HMI.sYELLOW; GVL_HMI.StatusHMI.sBannerTextColor := GVL_HMI.sBLACK;
    E_MachineState.ReadyToStart: GVL_HMI.StatusHMI.sMachineStatusText := 'SYSTEM READY TO START'; GVL_HMI.StatusHMI.sBannerBckColor := GVL_HMI.sGREEN; GVL_HMI.StatusHMI.sBannerTextColor := GVL_HMI.sWHITE;
    E_MachineState.AutoCycle: GVL_HMI.StatusHMI.sMachineStatusText := 'SYSTEM AUTO CYCLE'; GVL_HMI.StatusHMI.sBannerBckColor := GVL_HMI.sGREEN; GVL_HMI.StatusHMI.sBannerTextColor := GVL_HMI.sWHITE;
    E_MachineState.Stopping: GVL_HMI.StatusHMI.sMachineStatusText := 'STOPPING'; GVL_HMI.StatusHMI.sBannerBckColor := GVL_HMI.sGREY; GVL_HMI.StatusHMI.sBannerTextColor := GVL_HMI.sWHITE;
    E_MachineState.Stopped: GVL_HMI.StatusHMI.sMachineStatusText := 'CYCLE STOPPED'; GVL_HMI.StatusHMI.sBannerBckColor := GVL_HMI.sGREY; GVL_HMI.StatusHMI.sBannerTextColor := GVL_HMI.sWHITE;
    E_MachineState.Fault: GVL_HMI.StatusHMI.sMachineStatusText := 'IMMEDIATE FAULT'; GVL_HMI.StatusHMI.sBannerBckColor := GVL_HMI.sREDFail; GVL_HMI.StatusHMI.sBannerTextColor := GVL_HMI.sWHITE;
    E_MachineState.Manual: GVL_HMI.StatusHMI.sMachineStatusText := 'MANUAL MODE'; GVL_HMI.StatusHMI.sBannerBckColor := GVL_HMI.sBLUEInProgress; GVL_HMI.StatusHMI.sBannerTextColor := GVL_HMI.sWHITE;
END_CASE

END_PROGRAM

// ---- POUs/00_Application/PRG_WriteOutputs.TcPOU
PROGRAM PRG_WriteOutputs
VAR
END_VAR

GVL_IO.stOutputs.bSafetyRunRequest := GVL_MASTER.stOutputs.bSafetyRunRequest;
GVL_IO.stOutputs.bSafetyResetRequest := GVL_MASTER.stOutputs.bSafetyResetRequest;
GVL_IO.stOutputs.bSafetyErrorAcknowledgementRequest := GVL_MASTER.stOutputs.bSafetyErrorAcknowledgementRequest;
GVL_IO.stOutputs.bAirSupplyEnable := GVL_MASTER.stOutputs.bAirSupplyEnable;
GVL_IO.stOutputs.bMainDoorLockRequest := GVL_MASTER.stOutputs.bMainDoorLockRequest;
GVL_IO.stOutputs.bIndexRotatePortA := GVL_MASTER.stOutputs.bIndexRotatePortA;
GVL_IO.stOutputs.bIndexStopPortB := GVL_MASTER.stOutputs.bIndexStopPortB;
GVL_IO.stOutputs.bLedStart := GVL_MASTER.stOutputs.bLedStart;
GVL_IO.stOutputs.bLedReset := GVL_MASTER.stOutputs.bLedReset;
GVL_IO.stOutputs.bStatusIndicator := GVL_MASTER.stOutputs.bLedPass OR GVL_MASTER.stOutputs.bLedFail;
GVL_IO.stOutputs.bInternalLight := GVL_MASTER.stOutputs.bInternalLight;
GVL_IO.stOutputs.bNestLight := GVL_MASTER.stOutputs.bNestLight;

END_PROGRAM

// ---- POUs/01_Core/Process/FB_ProcessCycle.TcPOU
FUNCTION_BLOCK FB_ProcessCycle
VAR
    // STATE MACHINE
    eState                     : E_CycleState := E_CycleState.Disabled;

    // REQUESTS AND STATUS
    stRequestsInternal         : ST_ProcessCycleRequests;
    stStatusInternal           : ST_ProcessCycleStatus;

    // EDGE DETECTION
    rtProcessCycleTrigger      : R_TRIG;

    // SIMULATED PROCESS STATIONS
    tonAssemblyProcess         : TON;
    tonSiliconeProcess         : TON;
	
	// Timeout
	tonProcessCycleTimeout 		: TON;
	tonAutoCycleIdleTimeout 	: TON;
	
	bStopPending 				: BOOL;
	
	bSiliconeProcessCompleteLatched : BOOL;
    bAssemblyProcessCompleteLatched : BOOL;
	
END_VAR

METHOD PUBLIC Cyclic
VAR_INPUT
    bEnable          : BOOL;
    bResetRequest    : BOOL;
    bStopRequest     : BOOL;
    tSequenceTimeout : TIME;

    stInputs         : ST_ProcessCycleInputs;

END_VAR

VAR_OUTPUT
    stRequests       : ST_ProcessCycleRequests;
    stStatus         : ST_ProcessCycleStatus;
END_VAR
// The Process Cycle coordinates objects.
// It does not operate physical outputs directly.


// =========================================================
// CYCLIC DEFAULTS
// =========================================================

// stRequestsInternal.bStartProcessStation 			:= FALSE;
// stRequestsInternal.bStopProcessStation 				:= FALSE;
// stRequestsInternal.bCaptureProcessResult 			:= FALSE;
// stRequestsInternal.bStoreProcessResult 				:= FALSE;

stRequestsInternal.bSiliconeSupportExtend 			:= FALSE;
stRequestsInternal.bSiliconeSupportRetract 			:= FALSE;
stRequestsInternal.bAssemblySupportExtend 			:= FALSE;
stRequestsInternal.bAssemblySupportRetract 			:= FALSE;

stRequestsInternal.bStartSiliconeProcess 			:= FALSE;
stRequestsInternal.bStopSiliconeProcess 			:= FALSE;
stRequestsInternal.bCaptureSiliconeResult 			:= FALSE;
stRequestsInternal.bStoreSiliconeResult 			:= FALSE;

stRequestsInternal.bStartAssemblyProcess 			:= FALSE;
stRequestsInternal.bStopAssemblyProcess 			:= FALSE;
stRequestsInternal.bCaptureAssemblyResult 			:= FALSE;
stRequestsInternal.bStoreAssemblyResult 			:= FALSE;

stRequestsInternal.bPrepareOperatorExchange 		:= FALSE;
stRequestsInternal.bConfirmOperatorExchange 		:= FALSE;

stRequestsInternal.bRequestIndex 					:= FALSE;
stRequestsInternal.bRequestIndexRecovery 			:= FALSE;
stRequestsInternal.bUpdateNestPositions 			:= FALSE;

stStatusInternal.bCompletePulse 					:= FALSE;

// =========================================================
// PROCESS TRIGGER EDGE DETECTION
// =========================================================

rtProcessCycleTrigger(
    CLK := stInputs.bTwoHandsSafe
);

// =========================================================
// TIMEOUTS
// =========================================================

tonProcessCycleTimeout(
    IN := eState <> E_CycleState.Disabled
        AND eState <> E_CycleState.Initialising
        AND eState <> E_CycleState.WaitingForProcessCycleTrigger
        AND eState <> E_CycleState.CycleComplete
        AND eState <> E_CycleState.ControlledStop
		AND eState <> E_CycleState.WaitingForOperatorExchange
        AND eState <> E_CycleState.Fault,
    PT := tSequenceTimeout
);

IF tonProcessCycleTimeout.Q THEN
	stStatusInternal.bTimeoutFault := TRUE;
    eState := E_CycleState.Fault;
END_IF


/// =========================================================
// GLOBAL STATE CONTROL
// =========================================================

IF bResetRequest THEN
    // A reset starts a new process-cycle context.
    bStopPending := FALSE;
    bSiliconeProcessCompleteLatched := FALSE;
    bAssemblyProcessCompleteLatched := FALSE;
    stStatusInternal.bTimeoutFault := FALSE;
    eState := E_CycleState.Initialising;

ELSIF NOT bEnable THEN
    // No Stop request may remain stored while the
    // Process Cycle is disabled.
    bStopPending := FALSE;
    eState := E_CycleState.Disabled;

END_IF

// =========================================================
// STOP REQUEST LATCH
// ========================================================

// Memorise Stop only while the Process Cycle is enabled.
// The request remains stored until the current process and
// operator disposition have completed.
IF bEnable
    AND NOT bResetRequest AND bStopRequest THEN
    bStopPending := TRUE;
END_IF

// =========================================================
// PROCESS CYCLE STATE MACHINE
// =========================================================

CASE eState OF

    // -----------------------------------------------------
    // DISABLED
    // -----------------------------------------------------

    E_CycleState.Disabled:

        stStatusInternal.eMessage :=
            E_ProcessCycleMessage.None;

        IF bEnable THEN

            eState :=
                E_CycleState.Initialising;

        END_IF


    // -----------------------------------------------------
    // INITIALISING
    // -----------------------------------------------------

    E_CycleState.Initialising:

        stStatusInternal.eMessage :=
            E_ProcessCycleMessage.InitialisingProcessCycle;

        IF bEnable
            AND stInputs.bSafetyOk
            AND stInputs.bIndexReady
            AND stInputs.bIndexLocked
            AND stInputs.bSiliconeSupportRetracted
            AND stInputs.bAssemblySupportRetracted
        THEN

            eState :=
                E_CycleState.WaitingForProcessCycleTrigger;

        END_IF


    // -----------------------------------------------------
    // WAITING FOR PROCESS CYCLE TRIGGER
    // -----------------------------------------------------

   E_CycleState.WaitingForProcessCycleTrigger:

		stStatusInternal.eMessage := E_ProcessCycleMessage.WaitingForProcessCycleTrigger;
		// -----------------------------------------------------
		// SAFE STOP POINT
		// -----------------------------------------------------
		// No automatic process is active at this point.
		// A pending Stop request may therefore be executed
		// immediately without starting another cycle.
		IF bStopPending THEN
	
			bStopPending := FALSE;
			eState := E_CycleState.ControlledStop;
	
		ELSIF stInputs.bIndexFaulted
			OR stInputs.bSiliconeSupportFaulted
			OR stInputs.bAssemblySupportFaulted
		THEN
			eState := E_CycleState.Fault;
	
		ELSIF rtProcessCycleTrigger.Q
			AND stInputs.bSafetyOk
			AND stInputs.bIndexMoveAllowed
			AND stInputs.bIndexReady
			//AND stInputs.bIndexLocked
			AND stInputs.bSiliconeSupportRetracted
			AND stInputs.bAssemblySupportRetracted
		THEN
			eState := E_CycleState.ValidatingIndexPermissives;
		END_IF
		
		// -----------------------------------------------------
		// PREPARING OPERATOR EXCHANGE
		// -----------------------------------------------------
		
	E_CycleState.PreparingOperatorExchange:
		
			stStatusInternal.eMessage :=
				E_ProcessCycleMessage.PreparingOperatorExchange;
		
			stRequestsInternal.bPrepareOperatorExchange := TRUE;
		
			eState :=
				E_CycleState.WaitingForOperatorExchange;
		// -----------------------------------------------------
		// WAITING FOR OPERATOR EXCHANGE
		// -----------------------------------------------------
		
	E_CycleState.WaitingForOperatorExchange:
		
			stStatusInternal.eMessage :=
				E_ProcessCycleMessage.WaitingOperatorExchange;
	
		
			IF stInputs.bOperatorExchangeComplete THEN
		
				eState :=
					E_CycleState.ConfirmingOperatorExchange;
		
			END_IF

	// -----------------------------------------------------
	// CONFIRMING OPERATOR EXCHANGE
	// -----------------------------------------------------
	
	E_CycleState.ConfirmingOperatorExchange:
	
		stStatusInternal.eMessage := E_ProcessCycleMessage.ConfirmingOperatorExchange;
		stRequestsInternal.bConfirmOperatorExchange := TRUE;
		// -----------------------------------------------------
		// EXECUTE PENDING STOP
		// -----------------------------------------------------
		// The automatic cycle and operator disposition are
		// complete. A pending Stop request may now be executed.
		IF bStopPending THEN
	
			bStopPending := FALSE;
			eState := E_CycleState.ControlledStop;
		ELSE
			eState := E_CycleState.WaitingForProcessCycleTrigger;
		END_IF
    // -----------------------------------------------------
    // VALIDATING INDEX PERMISSIVES
    // -----------------------------------------------------

    E_CycleState.ValidatingIndexPermissives:

        stStatusInternal.eMessage := E_ProcessCycleMessage.ValidatingIndexPermissives;
		
        IF stInputs.bIndexFaulted THEN
            eState :=E_CycleState.Fault;

        ELSIF stInputs.bIndexMoveAllowed
            AND stInputs.bIndexReady
            AND stInputs.bIndexLocked
            AND stInputs.bSiliconeSupportRetracted
            AND stInputs.bAssemblySupportRetracted
        THEN

            eState :=
                E_CycleState.RequestingIndexMove;

        END_IF


    // -----------------------------------------------------
    // REQUESTING INDEX MOVE
    // -----------------------------------------------------

    E_CycleState.RequestingIndexMove:

        stRequestsInternal.bRequestIndex := TRUE;

        stStatusInternal.eMessage :=
            E_ProcessCycleMessage.RequestingIndexMove;

        IF stInputs.bIndexRequestAccepted THEN

            eState :=
                E_CycleState.WaitingForIndexStart;

        END_IF


    // -----------------------------------------------------
    // WAITING FOR INDEX START
    // -----------------------------------------------------

    E_CycleState.WaitingForIndexStart:

        stStatusInternal.eMessage :=
            E_ProcessCycleMessage.WaitingForIndexStart;

        IF stInputs.bIndexFaulted THEN

            eState :=
                E_CycleState.Fault;

        ELSIF stInputs.bIndexBusy
            OR stInputs.bIndexDone
        THEN

            eState :=
                E_CycleState.WaitingForIndexComplete;

        END_IF


    // -----------------------------------------------------
    // WAITING FOR INDEX COMPLETE
    // -----------------------------------------------------

    E_CycleState.WaitingForIndexComplete:

        stStatusInternal.eMessage :=E_ProcessCycleMessage.WaitingForIndexComplete;

       IF stInputs.bIndexFaulted THEN
			eState := E_CycleState.Fault;
		
		ELSIF stInputs.bIndexDone THEN
		
			IF stInputs.bIndexSamePositionDetected THEN
				stStatusInternal.eMessage := E_ProcessCycleMessage.IndexSamePositionDetected;
				eState := E_CycleState.CycleComplete;
		
			ELSIF stInputs.bSiliconeProcessRequired
				OR stInputs.bAssemblyProcessRequired
			THEN
				eState := E_CycleState.RequestingSupportsExtend;
		
			ELSE
				eState := E_CycleState.CycleComplete;
			END_IF
		
		END_IF


    // -----------------------------------------------------
    // REQUESTING SUPPORTS EXTEND
    // -----------------------------------------------------

    E_CycleState.RequestingSupportsExtend:

        stRequestsInternal.bSiliconeSupportExtend := stInputs.bSiliconeProcessRequired;
		stRequestsInternal.bAssemblySupportExtend := FALSE;

        stStatusInternal.eMessage :=
            E_ProcessCycleMessage.RequestingSupportsExtend;

        eState :=
            E_CycleState.WaitingForSupportsExtended;


    // -----------------------------------------------------
    // WAITING FOR SUPPORTS EXTENDED
    // -----------------------------------------------------

    E_CycleState.WaitingForSupportsExtended:

		stRequestsInternal.bSiliconeSupportExtend := stInputs.bSiliconeProcessRequired;
		stRequestsInternal.bAssemblySupportExtend := FALSE;
	
		stStatusInternal.eMessage :=
			E_ProcessCycleMessage.WaitingForSupportsExtended;
	
		IF (stInputs.bSiliconeProcessRequired AND stInputs.bSiliconeSupportFaulted)
			OR (stInputs.bAssemblyProcessRequired AND stInputs.bAssemblySupportFaulted)
		THEN
			eState := E_CycleState.Fault;
	
		ELSIF NOT stInputs.bSiliconeProcessRequired
			OR stInputs.bSiliconeSupportExtended
		THEN
			eState := E_CycleState.PreparingProcessStations;
		END_IF


    // -----------------------------------------------------
    // PREPARING PROCESS STATIONS
    // -----------------------------------------------------

    E_CycleState.PreparingProcessStations:

        stStatusInternal.eMessage :=
            E_ProcessCycleMessage.PreparingProcessStation;

        eState :=
            E_CycleState.StartingProcesses;


    // -----------------------------------------------------
	// STARTING PROCESSES
	// -----------------------------------------------------

	E_CycleState.StartingProcesses:
	
		stStatusInternal.eMessage := E_ProcessCycleMessage.StartingProcessEquipment;
			
		// Reset completion memory for the new process cycle.
		bSiliconeProcessCompleteLatched := FALSE;
		bAssemblyProcessCompleteLatched := FALSE;
	
		// Start only the processes required at the current
		// table positions.
		stRequestsInternal.bStartSiliconeProcess :=
			stInputs.bSiliconeProcessRequired;
	
		stRequestsInternal.bStartAssemblyProcess :=
			stInputs.bAssemblyProcessRequired;
	
		eState :=
			E_CycleState.WaitingForProcessesRunning;


	 // -----------------------------------------------------
	// WAITING FOR PROCESSES RUNNING
	// -----------------------------------------------------
	
	E_CycleState.WaitingForProcessesRunning:
	
	    // Raise Assembly Support only after the flipping station
    	// has reached the physical 0 degree position.
    	stRequestsInternal.bAssemblySupportExtend :=
        stInputs.bAssemblyProcessRequired
        AND
        (
            stInputs.bAssemblyAtZeroPosition
            OR stInputs.bAssemblySupportExtended
        );

		IF stInputs.bSiliconeProcessRequired
			AND stInputs.bSiliconeProcessComplete
		THEN
			bSiliconeProcessCompleteLatched := TRUE;
		END_IF
		
		IF stInputs.bAssemblyProcessRequired
			AND stInputs.bAssemblyProcessComplete
		THEN
			bAssemblyProcessCompleteLatched := TRUE;
		END_IF
	
		stStatusInternal.eMessage :=
			E_ProcessCycleMessage.StartingProcessEquipment;
	
		// Process equipment fault
		IF (stInputs.bSiliconeProcessRequired
				AND stInputs.bSiliconeProcessFaulted)
			OR
		   (stInputs.bAssemblyProcessRequired
				AND stInputs.bAssemblyProcessFaulted)
		THEN
	
			eState :=
				E_CycleState.Fault;
	
		// All required processes have started
		ELSIF
			(NOT stInputs.bSiliconeProcessRequired
				OR stInputs.bSiliconeProcessBusy
				OR bSiliconeProcessCompleteLatched)
			AND
			(NOT stInputs.bAssemblyProcessRequired
				OR stInputs.bAssemblyProcessBusy
				OR bAssemblyProcessCompleteLatched)
		THEN
	
			eState :=
				E_CycleState.WaitingForProcessesComplete;
	
		END_IF


    // -----------------------------------------------------
	// WAITING FOR PROCESSES COMPLETE
	// -----------------------------------------------------
	
	E_CycleState.WaitingForProcessesComplete:
		
			stRequestsInternal.bAssemblySupportExtend :=
		stInputs.bAssemblyProcessRequired
		AND
		(
			stInputs.bAssemblyAtZeroPosition
			OR stInputs.bAssemblySupportExtended
		);
	
		stStatusInternal.eMessage :=
			E_ProcessCycleMessage.WaitingForProcessesComplete;
			
		// Latch process completion.
		// Each process may complete at a different time and may be
		// reset by the machine coordinator after its result is stored.
		IF stInputs.bSiliconeProcessRequired AND stInputs.bSiliconeProcessComplete THEN
			bSiliconeProcessCompleteLatched := TRUE;
		END_IF
	
		IF stInputs.bAssemblyProcessRequired AND stInputs.bAssemblyProcessComplete THEN
			bAssemblyProcessCompleteLatched := TRUE;
		END_IF
	
		// Process fault
		IF (stInputs.bSiliconeProcessRequired
				AND stInputs.bSiliconeProcessFaulted)
			OR
		   (stInputs.bAssemblyProcessRequired
				AND stInputs.bAssemblyProcessFaulted)
		THEN
	
			eState :=
				E_CycleState.Fault;
	
		// All required processes completed
		ELSIF
			(NOT stInputs.bSiliconeProcessRequired
				OR bSiliconeProcessCompleteLatched)
			AND
			(NOT stInputs.bAssemblyProcessRequired
				OR bAssemblyProcessCompleteLatched)
		THEN
	
			eState :=
				E_CycleState.RequestingSupportsRetract;
	
		END_IF

    // -----------------------------------------------------
    // REQUESTING SUPPORTS RETRACT
    // -----------------------------------------------------

    E_CycleState.RequestingSupportsRetract:

        stRequestsInternal.bSiliconeSupportRetract := NOT stInputs.bSiliconeSupportRetracted;
		stRequestsInternal.bAssemblySupportRetract := NOT stInputs.bAssemblySupportRetracted;

        stStatusInternal.eMessage :=
            E_ProcessCycleMessage.RequestingSupportsRetract;

        eState :=
            E_CycleState.WaitingForSupportsRetracted;


    // -----------------------------------------------------
    // WAITING FOR SUPPORTS RETRACTED
    // -----------------------------------------------------

    E_CycleState.WaitingForSupportsRetracted:

        stRequestsInternal.bSiliconeSupportRetract := NOT stInputs.bSiliconeSupportRetracted;
		stRequestsInternal.bAssemblySupportRetract := NOT stInputs.bAssemblySupportRetracted;

        stStatusInternal.eMessage :=
            E_ProcessCycleMessage.WaitingForSupportsRetracted;

        IF (stInputs.bSiliconeProcessRequired AND stInputs.bSiliconeSupportFaulted)
			OR (stInputs.bAssemblyProcessRequired AND stInputs.bAssemblySupportFaulted)
		THEN
		
			eState := E_CycleState.Fault;
		
		ELSIF (NOT stInputs.bSiliconeProcessRequired OR stInputs.bSiliconeSupportRetracted)
			AND (NOT stInputs.bAssemblyProcessRequired OR stInputs.bAssemblySupportRetracted) 
			AND stInputs.bIndexMoveAllowed
		THEN
		
			eState := E_CycleState.CycleComplete;
		
		END_IF


    // -----------------------------------------------------
    // CYCLE COMPLETE
    // -----------------------------------------------------

    E_CycleState.CycleComplete:

        stStatusInternal.bCompletePulse := TRUE;

        stStatusInternal.eMessage :=
            E_ProcessCycleMessage.ProcessCycleComplete;

        eState :=
    		E_CycleState.PreparingOperatorExchange;


    // -----------------------------------------------------
	// CONTROLLED STOP
	// -----------------------------------------------------
	
	E_CycleState.ControlledStop:
	
		// Stop both station processes.
		stRequestsInternal.bStopSiliconeProcess := TRUE;
		stRequestsInternal.bStopAssemblyProcess := TRUE;
	
		// Retract supports only after their respective process has stopped.
        // This prevents the Silicone Support from moving away while the IVEK
        // dispense sequence is still active.
		stRequestsInternal.bSiliconeSupportRetract := NOT stInputs.bSiliconeProcessBusy;

        // Keep the Assembly Support in position until the flipping station has
        // completed its controlled return to home.
		stRequestsInternal.bAssemblySupportRetract := NOT stInputs.bAssemblyProcessBusy;
	
		stStatusInternal.eMessage :=
			E_ProcessCycleMessage.ControlledStopping;
	
		// Controlled stop is complete only when:
		// - Index is stopped
		// - Silicone process is not running
		// - Assembly process is not running
		// - Both supports are retracted
		IF NOT stInputs.bIndexBusy
			AND NOT stInputs.bSiliconeProcessBusy
			AND NOT stInputs.bAssemblyProcessBusy
			AND stInputs.bSiliconeSupportRetracted
			AND stInputs.bAssemblySupportRetracted
		THEN
	
			eState :=
				E_CycleState.Disabled;
	
		END_IF

    // -----------------------------------------------------
    // FAULT
    // -----------------------------------------------------
	
	E_CycleState.Fault:
	
		// Stop both station processes.
		stRequestsInternal.bStopSiliconeProcess := TRUE;
		stRequestsInternal.bStopAssemblyProcess := TRUE;
	
		stStatusInternal.eMessage :=
			E_ProcessCycleMessage.ProcessCycleFault;

END_CASE


// =========================================================
// STATUS MAPPING
// =========================================================

stStatusInternal.eState :=
    eState;

stStatusInternal.bActive :=
    bEnable
    AND eState <> E_CycleState.Disabled;

stStatusInternal.bIdle :=
    eState = E_CycleState.WaitingForProcessCycleTrigger;

stStatusInternal.bFaulted :=
    eState = E_CycleState.Fault;

stStatusInternal.bWaitingForPart :=
    FALSE;

stStatusInternal.bWaitingForOperator :=
    FALSE;

stStatusInternal.bWaitingForIndex :=
    eState = E_CycleState.ValidatingIndexPermissives
    OR eState = E_CycleState.RequestingIndexMove
    OR eState = E_CycleState.WaitingForIndexStart
    OR eState = E_CycleState.WaitingForIndexComplete;

stStatusInternal.bWaitingForSupports :=
    eState = E_CycleState.RequestingSupportsExtend
    OR eState = E_CycleState.WaitingForSupportsExtended
    OR eState = E_CycleState.RequestingSupportsRetract
    OR eState = E_CycleState.WaitingForSupportsRetracted;

stStatusInternal.bSiliconeSupportExtended :=
    stInputs.bSiliconeSupportExtended;

stStatusInternal.bSiliconeSupportRetracted :=
    stInputs.bSiliconeSupportRetracted;

stStatusInternal.bAssemblySupportExtended :=
    stInputs.bAssemblySupportExtended;

stStatusInternal.bAssemblySupportRetracted :=
    stInputs.bAssemblySupportRetracted;

// =========================================================
// PROCESS STATUS
// =========================================================

stStatusInternal.bSiliconeProcessRunning :=
    stInputs.bSiliconeProcessRequired
    AND stInputs.bSiliconeProcessBusy;

stStatusInternal.bSiliconeProcessComplete :=
    NOT stInputs.bSiliconeProcessRequired
    OR stInputs.bSiliconeProcessComplete;


stStatusInternal.bAssemblyProcessRunning :=
    stInputs.bAssemblyProcessRequired
    AND stInputs.bAssemblyProcessBusy;

stStatusInternal.bAssemblyProcessComplete :=
    NOT stInputs.bAssemblyProcessRequired
    OR stInputs.bAssemblyProcessComplete;
// =========================================================
// MESSAGE MAPPING
// =========================================================

CASE stStatusInternal.eMessage OF

    E_ProcessCycleMessage.None:
        stStatusInternal.sMessage := '';
	
	E_ProcessCycleMessage.IndexSamePositionDetected:
    stStatusInternal.sMessage :=
        'Index returned to the same position - press and hold the two-hand controls to retry';

    E_ProcessCycleMessage.InitialisingProcessCycle:
        stStatusInternal.sMessage := 'Initialising automatic process cycle';

    E_ProcessCycleMessage.WaitingForProcessCycleTrigger:
        stStatusInternal.sMessage := 'Place both hands on the two-hand controls to start the cycle';

    E_ProcessCycleMessage.ValidatingIndexPermissives:
        stStatusInternal.sMessage := 'Validating index movement conditions';

    E_ProcessCycleMessage.RequestingIndexMove:
        stStatusInternal.sMessage := 'Requesting index table movement';

    E_ProcessCycleMessage.WaitingForIndexStart:
        stStatusInternal.sMessage := 'Waiting for index table movement to start';

    E_ProcessCycleMessage.WaitingForIndexComplete:
        stStatusInternal.sMessage := 'Index table moving';

    E_ProcessCycleMessage.RequestingSupportsExtend:
        stStatusInternal.sMessage := 'Requesting support extension';

    E_ProcessCycleMessage.WaitingForSupportsExtended:
        stStatusInternal.sMessage := 'Waiting for Silicone and Assembly Supports to extend';

    E_ProcessCycleMessage.PreparingProcessStation:
        stStatusInternal.sMessage := 'Preparing Assembly and Silicone processes';

    E_ProcessCycleMessage.StartingProcessEquipment:
        stStatusInternal.sMessage := 'Starting Assembly and Silicone processes';

    E_ProcessCycleMessage.WaitingForProcessesComplete:
        //stStatusInternal.sMessage := 'Assembly and Silicone processes in progress';
		IF stInputs.bSiliconeProcessRequired AND stInputs.bAssemblyProcessRequired THEN
			
			stStatusInternal.sMessage := 'Assembly and Silicone processes in progress';
	
		ELSIF stInputs.bSiliconeProcessRequired THEN
	
			stStatusInternal.sMessage := 'Silicone in progress';
	
		ELSIF stInputs.bAssemblyProcessRequired THEN
	
			stStatusInternal.sMessage := 'Assembly in progress';
	
		ELSE
	
			stStatusInternal.sMessage := 'Processes in progress';
	
		END_IF

    E_ProcessCycleMessage.RequestingSupportsRetract:
        stStatusInternal.sMessage := 'Requesting support retraction';

    E_ProcessCycleMessage.WaitingForSupportsRetracted:
        stStatusInternal.sMessage := 'Waiting for Silicone and Assembly Supports to retract';

    E_ProcessCycleMessage.ProcessCycleComplete:
        stStatusInternal.sMessage := 'Automatic process cycle complete';

    E_ProcessCycleMessage.ControlledStopping:
        stStatusInternal.sMessage := 'Stopping automatic cycle safely';

    E_ProcessCycleMessage.ProcessCycleFault:
        stStatusInternal.sMessage := 'Automatic process cycle fault';

ELSE

    stStatusInternal.sMessage := '';

END_CASE



// =========================================================
// OUTPUT PUBLICATION
// =========================================================

stRequests :=
    stRequestsInternal;

stStatus :=
    stStatusInternal;
END_METHOD

METHOD PUBLIC Initialise
eState := E_CycleState.Disabled;

bStopPending := FALSE;
bSiliconeProcessCompleteLatched := FALSE;
bAssemblyProcessCompleteLatched := FALSE;

stRequestsInternal.bPrepareOperatorExchange := FALSE;
stRequestsInternal.bConfirmOperatorExchange := FALSE;
stRequestsInternal.bRequestIndex := FALSE;
stRequestsInternal.bRequestIndexRecovery := FALSE;
stRequestsInternal.bUpdateNestPositions := FALSE;
stStatusInternal.bCompletePulse := FALSE;
stStatusInternal.bFaulted := FALSE;
stStatusInternal.bTimeoutFault := FALSE;
stStatusInternal.eMessage := E_ProcessCycleMessage.None;
END_METHOD

END_FUNCTION_BLOCK

// ---- POUs/01_Core/Process/FB_ProcessStation.TcPOU
FUNCTION_BLOCK FB_ProcessStation
VAR
    ipEquipment       : I_ProcessEquipment;
    bConfigured       : BOOL;
    eState            : E_ProcessStationState := E_ProcessStationState.Disabled;
    eFault            : E_ProcessStationFault := E_ProcessStationFault.None;
    stResult          : ST_ProcessResult;
    stStatusInternal  : ST_ProcessStationStatus;
    tonCylinder       : TON;
    tonProcess        : TON;
END_VAR

METHOD PUBLIC Configure : BOOL
VAR_INPUT
 ipNewEquipment : I_ProcessEquipment;
END_VAR
ipEquipment := ipNewEquipment;
bConfigured := TRUE;
Configure := TRUE;
END_METHOD

METHOD PUBLIC Cyclic : BOOL
VAR_INPUT
    bEnable                  : BOOL;
    bAutomaticStartRequest   : BOOL;
    bManualEnable            : BOOL;
    bManualExtendRequest     : BOOL;
    bManualRetractRequest    : BOOL;
    bStopRequest             : BOOL;
    bResetRequest            : BOOL;
    bPartPresent             : BOOL;
    bProcessPermissive       : BOOL;
    bIndexReady              : BOOL;
    bIndexLocked             : BOOL;
    bIndexBusy               : BOOL;
    bProcessSafetyPermitted  : BOOL;
    bMainDoorSafe            : BOOL;
    bCylinderExtended        : BOOL;
    bCylinderRetracted       : BOOL;
    tCylinderTimeout         : TIME;
    tProcessTimeout          : TIME;
	bAirSupplySafe 			 : BOOL;
	
END_VAR
VAR_OUTPUT
    bCylinderExtendOutput    : BOOL;
    bCylinderRetractOutput   : BOOL;
END_VAR
bCylinderExtendOutput := FALSE;
bCylinderRetractOutput := FALSE;

IF bConfigured THEN
    ipEquipment.Cyclic();
END_IF

stStatusInternal.bExtendPermissive :=
    bProcessSafetyPermitted
    AND bMainDoorSafe
    AND bIndexReady
    AND bIndexLocked
	AND bAirSupplySafe
    AND NOT bIndexBusy;
	
stStatusInternal.bRetractPermissive :=
    bProcessSafetyPermitted
    AND bAirSupplySafe
    AND NOT bIndexBusy;

IF bCylinderExtended AND bCylinderRetracted THEN
    eFault := E_ProcessStationFault.CylinderSensorMismatch;
    eState := E_ProcessStationState.Fault;
END_IF

// =========================================================
// RESET
// =========================================================
//
// Reset clears the Process Station fault only after the
// contradictory cylinder-sensor condition has disappeared.
//
// Pneumatic position recovery is NOT performed during Fault.
// The station returns to Disabled and will recover its safe
// position when it is enabled again during Initialising.
// =========================================================

IF bResetRequest THEN

    IF bConfigured THEN
        ipEquipment.RequestReset();
    END_IF

    // A simultaneous Extended + Retracted indication is a real
    // sensor contradiction and must not be cleared by Reset.
    IF NOT (bCylinderExtended AND bCylinderRetracted) THEN

        eFault := E_ProcessStationFault.None;
        stResult.bValid := FALSE;

        eState := E_ProcessStationState.Disabled;

    END_IF

END_IF

// =========================================================
// GLOBAL CONTROL
// =========================================================

IF NOT bConfigured THEN

    eFault := E_ProcessStationFault.EquipmentFault;
    eState := E_ProcessStationState.Fault;


ELSIF bStopRequest THEN

    // Fault / Stopping:
    //
    // Stop the process equipment, but do not attempt pneumatic
    // recovery here. The machine air supply may already have
    // been removed.
    ipEquipment.RequestStop();

    IF eState <> E_ProcessStationState.Fault THEN
        eState := E_ProcessStationState.Disabled;
    END_IF


ELSIF bManualEnable THEN

    ipEquipment.RequestStop();
    eState := E_ProcessStationState.Disabled;


ELSIF NOT bEnable THEN

    // Station disabled outside Automatic / Initialising.
    //
    // Do not start a retract sequence here because air may not
    // currently be available.
    ipEquipment.RequestStop();

    eState := E_ProcessStationState.Disabled;

END_IF

CASE eState OF
	
    E_ProcessStationState.Disabled:

    // Recovery is only performed when the station is enabled.
    // Machine Initialising enables the station after requesting
    // the pneumatic supply.
    IF bEnable THEN
        IF bCylinderRetracted THEN
            eState := E_ProcessStationState.Idle;
        ELSIF stStatusInternal.bRetractPermissive THEN
            //eState := E_ProcessStationState.Retracting;
        END_IF
    END_IF

    E_ProcessStationState.Idle:
        bCylinderRetractOutput := NOT bCylinderRetracted;
        IF bManualEnable THEN
            IF bManualExtendRequest AND bManualRetractRequest THEN
                eFault := E_ProcessStationFault.CommandConflict;
                eState := E_ProcessStationState.Fault;
            ELSIF bManualExtendRequest AND stStatusInternal.bExtendPermissive THEN
                eState := E_ProcessStationState.Advancing;
            ELSIF bManualRetractRequest THEN
                eState := E_ProcessStationState.Retracting;
            END_IF
        ELSIF bEnable AND bAutomaticStartRequest AND bPartPresent AND bProcessPermissive AND ipEquipment.IsReady() THEN
            stResult.bValid := FALSE;
            eState := E_ProcessStationState.Advancing;
        END_IF

    E_ProcessStationState.Advancing:
        IF NOT stStatusInternal.bExtendPermissive THEN
            eFault := E_ProcessStationFault.SafetyLostDuringMovement;
            eState := E_ProcessStationState.Fault;
        ELSE
            bCylinderExtendOutput := NOT bCylinderExtended;
            IF bCylinderExtended THEN
                IF bManualEnable THEN eState := E_ProcessStationState.Advanced; ELSE eState := E_ProcessStationState.StartingEquipment; END_IF
            END_IF
        END_IF

    E_ProcessStationState.Advanced:
        IF bManualRetractRequest OR NOT bManualEnable THEN eState := E_ProcessStationState.Retracting; END_IF

    E_ProcessStationState.StartingEquipment:
        IF NOT bCylinderExtended OR NOT bIndexReady OR NOT bIndexLocked THEN
            eFault := E_ProcessStationFault.IndexNotLocked;
            eState := E_ProcessStationState.Fault;
        ELSIF ipEquipment.RequestStart() THEN
            eState := E_ProcessStationState.Processing;
        ELSIF ipEquipment.IsFaulted() THEN
            eFault := E_ProcessStationFault.EquipmentFault;
            eState := E_ProcessStationState.Fault;
        END_IF

    E_ProcessStationState.Processing:
        bCylinderExtendOutput := TRUE;
        IF ipEquipment.IsDone() THEN
            stResult := ipEquipment.GetResult();
            eState := E_ProcessStationState.StoppingEquipment;
        ELSIF ipEquipment.IsFaulted() THEN
            stResult := ipEquipment.GetResult();
            eFault := E_ProcessStationFault.EquipmentFault;
            eState := E_ProcessStationState.Fault;
        END_IF

    E_ProcessStationState.StoppingEquipment:
        ipEquipment.RequestStop();
        IF NOT ipEquipment.IsBusy() THEN eState := E_ProcessStationState.Retracting; END_IF

    E_ProcessStationState.Retracting:
        bCylinderRetractOutput := NOT bCylinderRetracted;
        IF bCylinderRetracted AND NOT ipEquipment.IsBusy() THEN
			
            IF stResult.bValid THEN 
				eState := E_ProcessStationState.Complete;
            ELSIF bEnable OR bManualEnable THEN 
				eState := E_ProcessStationState.Idle;
            ELSE 
				eState := E_ProcessStationState.Disabled;
            END_IF
			
        END_IF

    E_ProcessStationState.Complete:
        bCylinderRetractOutput := NOT bCylinderRetracted;
        IF bCylinderRetracted THEN
            IF bEnable OR bManualEnable THEN eState := E_ProcessStationState.Idle; ELSE eState := E_ProcessStationState.Disabled; END_IF
        END_IF

    E_ProcessStationState.Fault:

    // Fault is a non-recovery state.
    // Pneumatic recovery is performed during machine Initialising.
    ipEquipment.RequestStop();

    bCylinderExtendOutput := FALSE;
    bCylinderRetractOutput := FALSE;
END_CASE

tonCylinder(
    IN := ((eState = E_ProcessStationState.Advancing) AND NOT bCylinderExtended)
       OR ((eState = E_ProcessStationState.Retracting) AND NOT bCylinderRetracted),
    PT := tCylinderTimeout);
IF tonCylinder.Q THEN
    IF eState = E_ProcessStationState.Advancing THEN eFault := E_ProcessStationFault.CylinderExtendTimeout;
    ELSE eFault := E_ProcessStationFault.CylinderRetractTimeout;
    END_IF
    eState := E_ProcessStationState.Fault;
END_IF

tonProcess(IN := eState = E_ProcessStationState.Processing, PT := tProcessTimeout);
IF tonProcess.Q THEN
    ipEquipment.RequestStop();
    stResult.bValid := TRUE;
    stResult.bPassed := FALSE;
    stResult.eCode := E_ProcessResultCode.Timeout;
    eFault := E_ProcessStationFault.ProcessTimeout;
    eState := E_ProcessStationState.Fault;
END_IF

stStatusInternal.eState := eState;
stStatusInternal.eFault := eFault;
stStatusInternal.bReady := eState = E_ProcessStationState.Idle;
stStatusInternal.bBusy := (eState = E_ProcessStationState.Advancing) OR (eState = E_ProcessStationState.StartingEquipment) OR (eState = E_ProcessStationState.Processing) OR (eState = E_ProcessStationState.StoppingEquipment) OR (eState = E_ProcessStationState.Retracting);
stStatusInternal.bFaulted := eState = E_ProcessStationState.Fault;
stStatusInternal.bSafePosition := bCylinderRetracted AND NOT ipEquipment.IsBusy();
stStatusInternal.bCylinderExtended := bCylinderExtended;
stStatusInternal.bCylinderRetracted := bCylinderRetracted;
stStatusInternal.bAutomaticRequestActive := bEnable AND bAutomaticStartRequest;
stStatusInternal.bManualRequestActive := bManualEnable AND (bManualExtendRequest OR bManualRetractRequest);
stStatusInternal.bEquipmentReady := ipEquipment.IsReady();
stStatusInternal.bEquipmentBusy := ipEquipment.IsBusy();
stStatusInternal.bEquipmentFaulted := ipEquipment.IsFaulted();
CASE eState OF
    E_ProcessStationState.Disabled: stStatusInternal.sMessage := 'Process station disabled';
    E_ProcessStationState.Idle: stStatusInternal.sMessage := 'Process station ready';
    E_ProcessStationState.Advancing: stStatusInternal.sMessage := 'Advancing Silicone Support Cylinder';
    E_ProcessStationState.Advanced: stStatusInternal.sMessage := 'Silicone Support Cylinder extended';
    E_ProcessStationState.StartingEquipment: stStatusInternal.sMessage := 'Starting process equipment';
    E_ProcessStationState.Processing: stStatusInternal.sMessage := 'Process in progress';
    E_ProcessStationState.StoppingEquipment: stStatusInternal.sMessage := 'Stopping process equipment';
    E_ProcessStationState.Retracting: stStatusInternal.sMessage := 'Retracting Silicone Support Cylinder';
    E_ProcessStationState.Complete: stStatusInternal.sMessage := 'Process complete';
    E_ProcessStationState.Fault: stStatusInternal.sMessage := 'Process station fault';
END_CASE
Cyclic := NOT stStatusInternal.bFaulted;
END_METHOD

METHOD PUBLIC GetResult : ST_ProcessResult
GetResult := stResult;
END_METHOD

METHOD PUBLIC GetStatus : ST_ProcessStationStatus
GetStatus := stStatusInternal;
END_METHOD

METHOD PUBLIC IndexPermissive : BOOL
IndexPermissive := stStatusInternal.bSafePosition AND NOT stStatusInternal.bFaulted;
END_METHOD

METHOD PUBLIC Initialise
stResult.bValid := FALSE;
eFault := E_ProcessStationFault.None;
IF bConfigured THEN eState := E_ProcessStationState.Idle; ELSE eState := E_ProcessStationState.Disabled; END_IF
tonCylinder(IN := FALSE);
tonProcess(IN := FALSE);
END_METHOD

METHOD PUBLIC IsComplete : BOOL
IsComplete := stResult.bValid AND eState = E_ProcessStationState.Complete;
END_METHOD

METHOD PUBLIC IsFaulted : BOOL
IsFaulted := stStatusInternal.bFaulted;
END_METHOD

METHOD PUBLIC IsSafePosition : BOOL
IsSafePosition := stStatusInternal.bSafePosition;
END_METHOD

METHOD PUBLIC ResetFault : BOOL
VAR_INPUT
 bCylinderExtended : BOOL;
 bCylinderRetracted : BOOL;
END_VAR
ResetFault := FALSE;
IF NOT (bCylinderExtended AND bCylinderRetracted) THEN
 eFault := E_ProcessStationFault.None;
 eState := E_ProcessStationState.Retracting;
 ResetFault := TRUE;
END_IF
END_METHOD

END_FUNCTION_BLOCK

// ---- POUs/02_Components/Pneumatics/FB_PuckLocker.TcPOU
FUNCTION_BLOCK FB_PuckLocker
VAR
    eState                   : E_PuckLockerState := E_PuckLockerState.Disabled;
    stStatusInternal         : ST_PuckLockerStatus;
    bReleaseRequested        : BOOL;
    bPartRemoved             : BOOL;
    bPreviousPuckDetected    : BOOL;
    bAcknowledgePrevious     : BOOL;
    tonRemovalConfirm        : TON;
END_VAR

